(* IEC 61131-3 sources: llm-plc-st-eval/codesys, 25 files *)

(* ---- PRG_Test_A1.st ---- *)
(*
    BANCO DE PRUEBA AUTOVERIFICABLE - Tarea A1 (FB_PID con anti-windup por clamping)
    ---------------------------------------------------------------------------
    Validado en codesys/validar_harness_A1.py: 12 implementaciones (3 correctas,
    con integracion rectangular, integral previa y trapezoidal, y 9 defectuosas).
    Tabla generada desde el validador. tipo: 0 = valor +-tol, 1 = CV <= eVal,
    2 = CV >= eVal.

    TOLERANCIAS (aprobadas por Luis y su asesora, 30-09-2026):
  solo P: +-0.01 | integral: +-2 pasos de muestreo | derivada: +-5 % del termino
  derivativo | saturacion exacta (+-0.001) | anti-windup: sale de la saturacion en
  menos de 1 s tras invertir el error | sentido: PV < SP -> CV sube.

TIEMPO VIRTUAL: ciclo := T#100MS fijo; pasos por NUMERO DE LLAMADAS. Cada
escenario usa su PROPIA instancia del FB (fbP, fbI, fbD, fbW), para que el estado
interno de un escenario (p. ej. una integral acumulada) no contamine otro.

Paso  instancia  (Kp, Ti, Td, SP, PV) llamadas -> comprobacion
  0   fbP  (2, 0, 0, 50, 40)     5 -> CV = 20.0 +-0.01     solo P, sentido
  1   fbP  (2, 0, 0, 50, 60)     5 -> CV = 0.0 +-0.001     saturacion baja
  2   fbP  (2, 0, 0, 50,-20)     5 -> CV = 100.0 +-0.001   saturacion alta
  3   fbP  (2,-1, 0, 50, 45)     5 -> CV = 10.0 +-0.01     Ti < 0: sin integral
  4   fbI  (1,10, 0, 50, 45)   100 -> CV = 10.0 +-0.10     5 + 0.5*10 s
  5   fbI  (1,10, 0, 50, 45)   100 -> CV = 15.0 +-0.10     5 + 0.5*20 s
  6   fbD  (1, 0, 2, 50+0.1k, 40) 50 -> CV = 17.0 +-0.10   e = 15, Td*de/dt = 2 (SP en rampa:
                                                           la derivada sobre PV daria 0)
  7   fbW  (1, 5, 0,100,  0)   300 -> CV = 100.0 +-0.001   30 s saturado en alto
  8   fbW  (1, 5, 0,100,110)    10 -> CV <= 99.5            sale de 100 en < 1 s
  9   fbW  (1, 5, 0,  0,200)   300 -> CV = 0.0 +-0.001     30 s saturado en bajo
 10   fbW  (1, 5, 0,  0,-10)    10 -> CV >= 0.5             sale de 0 en < 1 s
*)
PROGRAM PRG_Test_A1
VAR CONSTANT
    ULTIMO_PASO : INT := 10;
END_VAR
VAR
    fbP, fbI, fbD, fbW : FB_PID;    (* una instancia por escenario *)
    ins        : INT;
    Kp, Ti, Td : REAL;
    SPbase, PV : REAL;
    rampa      : BOOL;
    kRampa     : INT;
    SP, CV     : REAL;
    nLlamadas, k, tipo : INT;
    eVal, tol  : REAL;
    bien       : BOOL;
    paso       : INT := 0;
    finalizado : BOOL;

    resultado : ARRAY[0..10] OF INT;
    nPasan    : INT;
    veredicto : INT := 0;
    i         : INT;
END_VAR

IF NOT finalizado THEN
    (* 1. Definicion del paso *)
    CASE paso OF
        0: ins := 0; Kp := 2.0; Ti := 0.0; Td := 0.0; SPbase := 50.0; rampa := FALSE; PV := 40.0; nLlamadas := 5; tipo := 0; eVal := 20.0; tol := 0.01;
        1: ins := 0; Kp := 2.0; Ti := 0.0; Td := 0.0; SPbase := 50.0; rampa := FALSE; PV := 60.0; nLlamadas := 5; tipo := 0; eVal := 0.0; tol := 0.001;
        2: ins := 0; Kp := 2.0; Ti := 0.0; Td := 0.0; SPbase := 50.0; rampa := FALSE; PV := -20.0; nLlamadas := 5; tipo := 0; eVal := 100.0; tol := 0.001;
        3: ins := 0; Kp := 2.0; Ti := -1.0; Td := 0.0; SPbase := 50.0; rampa := FALSE; PV := 45.0; nLlamadas := 5; tipo := 0; eVal := 10.0; tol := 0.01;
        4: ins := 1; Kp := 1.0; Ti := 10.0; Td := 0.0; SPbase := 50.0; rampa := FALSE; PV := 45.0; nLlamadas := 100; tipo := 0; eVal := 10.0; tol := 0.1;
        5: ins := 1; Kp := 1.0; Ti := 10.0; Td := 0.0; SPbase := 50.0; rampa := FALSE; PV := 45.0; nLlamadas := 100; tipo := 0; eVal := 15.0; tol := 0.1;
        6: ins := 2; Kp := 1.0; Ti := 0.0; Td := 2.0; SPbase := 50.0; rampa := TRUE; PV := 40.0; nLlamadas := 50; tipo := 0; eVal := 17.0; tol := 0.1;
        7: ins := 3; Kp := 1.0; Ti := 5.0; Td := 0.0; SPbase := 100.0; rampa := FALSE; PV := 0.0; nLlamadas := 300; tipo := 0; eVal := 100.0; tol := 0.001;
        8: ins := 3; Kp := 1.0; Ti := 5.0; Td := 0.0; SPbase := 100.0; rampa := FALSE; PV := 110.0; nLlamadas := 10; tipo := 1; eVal := 99.5; tol := 0.0;
        9: ins := 3; Kp := 1.0; Ti := 5.0; Td := 0.0; SPbase := 0.0; rampa := FALSE; PV := 200.0; nLlamadas := 300; tipo := 0; eVal := 0.0; tol := 0.001;
        10: ins := 3; Kp := 1.0; Ti := 5.0; Td := 0.0; SPbase := 0.0; rampa := FALSE; PV := -10.0; nLlamadas := 10; tipo := 2; eVal := 0.5; tol := 0.0;
    END_CASE

    (* 2. Consigna (en rampa en el escenario derivativo) *)
    IF rampa THEN
        kRampa := kRampa + 1;
        SP := SPbase + 0.1 * INT_TO_REAL(kRampa);
    ELSE
        SP := SPbase;
    END_IF

    (* 3. Una llamada por scan a la instancia del escenario, ciclo virtual 100 ms *)
    CASE ins OF
        0: fbP(SP := SP, PV := PV, Kp := Kp, Ti := Ti, Td := Td, ciclo := T#100MS); CV := fbP.CV;
        1: fbI(SP := SP, PV := PV, Kp := Kp, Ti := Ti, Td := Td, ciclo := T#100MS); CV := fbI.CV;
        2: fbD(SP := SP, PV := PV, Kp := Kp, Ti := Ti, Td := Td, ciclo := T#100MS); CV := fbD.CV;
        3: fbW(SP := SP, PV := PV, Kp := Kp, Ti := Ti, Td := Td, ciclo := T#100MS); CV := fbW.CV;
    END_CASE
    k := k + 1;

    (* 4. Evaluacion al completar las llamadas del paso *)
    IF k >= nLlamadas THEN
        CASE tipo OF
            0: bien := ABS(CV - eVal) <= tol;
            1: bien := CV <= eVal;
            2: bien := CV >= eVal;
        END_CASE
        IF bien THEN
            resultado[paso] := 1;
        ELSE
            resultado[paso] := 2;
        END_IF
        k := 0;
        IF paso < ULTIMO_PASO THEN
            paso := paso + 1;
        ELSE
            finalizado := TRUE;
        END_IF
    END_IF
END_IF

(* 5. Veredicto global *)
IF finalizado AND veredicto = 0 THEN
    nPasan := 0;
    FOR i := 0 TO ULTIMO_PASO DO
        IF resultado[i] = 1 THEN
            nPasan := nPasan + 1;
        END_IF
    END_FOR
    IF nPasan = (ULTIMO_PASO + 1) THEN
        veredicto := 1;
    ELSE
        veredicto := 2;
    END_IF
END_IF

(* ---- PRG_Test_A2.st ---- *)
(*
    BANCO DE PRUEBA AUTOVERIFICABLE - Tarea A2 (FB_Batch: receta por lotes de 5 fases)
    ---------------------------------------------------------------------------
    Validado en codesys/validar_harness_A2.py: 9 implementaciones (1 correcta y
    8 defectuosas), ciclos de 4, 10 y 20 ms. Tabla generada desde el validador.
    Al final de cada paso se exige la fase esperada y que este activa exactamente
    la salida de esa fase (fase 0: ninguna).

    Paso: (nA,nB,nVac,ini,abo,temp) duracion -> fase esperada
  0 (F,F,F,F,F,20)   0.2 s -> 0   reposo CON producto
  1 (F,F,F,F,T,20)   0.2 s -> 0   abort en reposo: sin efecto
  2 (F,F,F,T,F,20)   0.2 s -> 1   inicio
  3 (F,F,F,F,F,20)   0.2 s -> 1   espera nivelA
  4 (T,F,F,F,F,20)   0.2 s -> 2
  5 (T,F,F,T,F,20)   0.2 s -> 2   inicio durante la receta: se ignora
  6 (T,T,F,F,F,20)   0.2 s -> 3
  7 (T,T,F,F,F,59.9) 0.2 s -> 3   59.9 no basta
  8 (T,T,F,F,F,60.0) 0.2 s -> 4   60.0 o mas
  9 (T,T,F,F,F,60.0) 118  s -> 4   mezcla: aun no cumple 120 s
 10 (T,T,F,F,F,60.0) 3.0 s -> 5   ya cumplio
 11 (T,T,T,F,F,60.0) 0.2 s -> 0   vacio: reposo
 12 (F,F,F,T,F,20)   0.2 s -> 1   nueva receta (con producto)
 13 (F,F,F,F,T,20)   0.2 s -> 5   abort con producto: descarga
 14 (F,F,F,F,F,20)   0.2 s -> 5   sigue descargando
 15 (F,F,T,F,F,20)   0.2 s -> 0
 16 (F,F,T,T,F,20)   0.2 s -> 1   receta con reactor vacio
 17 (F,F,T,F,T,20)   0.2 s -> 0   abort sin producto: directo a reposo
 18 (F,F,F,T,F,20)   0.2 s -> 1
 19 (T,F,F,F,F,20)   0.2 s -> 2
 20 (T,T,F,F,F,20)   0.2 s -> 3   calentando
 21 (T,T,F,F,T,20)   0.2 s -> 5   abort en fase 3: calentador cerrado, descarga
 22 (T,T,F,F,F,20)   0.2 s -> 5
 23 (T,T,F,F,T,20)   0.2 s -> 5   abort durante la descarga: continua
 24 (T,T,T,F,F,20)   0.2 s -> 0
*)
PROGRAM PRG_Test_A2
VAR CONSTANT
    ULTIMO_PASO : INT := 24;
END_VAR
VAR
    fb : FB_Batch;                  (* bloque bajo prueba *)
    nivelA, nivelB, nivelVacio, btnInicio, btnAbort : BOOL;
    temp  : REAL;
    eFase : INT;
    salidasOk : BOOL;

    paso       : INT := 0;
    tEspera    : TIME;
    tPaso      : TON;
    pulsoReset : BOOL;
    finalizado : BOOL;

    resultado : ARRAY[0..24] OF INT;
    nPasan    : INT;
    veredicto : INT := 0;
    i         : INT;
END_VAR

(* 1. Entradas, duracion y fase esperada del paso *)
IF NOT finalizado THEN
    CASE paso OF
        0: nivelA := FALSE; nivelB := FALSE; nivelVacio := FALSE; btnInicio := FALSE; btnAbort := FALSE;
            temp := 20.0; tEspera := T#200MS; eFase := 0;
        1: nivelA := FALSE; nivelB := FALSE; nivelVacio := FALSE; btnInicio := FALSE; btnAbort := TRUE;
            temp := 20.0; tEspera := T#200MS; eFase := 0;
        2: nivelA := FALSE; nivelB := FALSE; nivelVacio := FALSE; btnInicio := TRUE; btnAbort := FALSE;
            temp := 20.0; tEspera := T#200MS; eFase := 1;
        3: nivelA := FALSE; nivelB := FALSE; nivelVacio := FALSE; btnInicio := FALSE; btnAbort := FALSE;
            temp := 20.0; tEspera := T#200MS; eFase := 1;
        4: nivelA := TRUE; nivelB := FALSE; nivelVacio := FALSE; btnInicio := FALSE; btnAbort := FALSE;
            temp := 20.0; tEspera := T#200MS; eFase := 2;
        5: nivelA := TRUE; nivelB := FALSE; nivelVacio := FALSE; btnInicio := TRUE; btnAbort := FALSE;
            temp := 20.0; tEspera := T#200MS; eFase := 2;
        6: nivelA := TRUE; nivelB := TRUE; nivelVacio := FALSE; btnInicio := FALSE; btnAbort := FALSE;
            temp := 20.0; tEspera := T#200MS; eFase := 3;
        7: nivelA := TRUE; nivelB := TRUE; nivelVacio := FALSE; btnInicio := FALSE; btnAbort := FALSE;
            temp := 59.9; tEspera := T#200MS; eFase := 3;
        8: nivelA := TRUE; nivelB := TRUE; nivelVacio := FALSE; btnInicio := FALSE; btnAbort := FALSE;
            temp := 60.0; tEspera := T#200MS; eFase := 4;
        9: nivelA := TRUE; nivelB := TRUE; nivelVacio := FALSE; btnInicio := FALSE; btnAbort := FALSE;
            temp := 60.0; tEspera := T#118000MS; eFase := 4;
        10: nivelA := TRUE; nivelB := TRUE; nivelVacio := FALSE; btnInicio := FALSE; btnAbort := FALSE;
            temp := 60.0; tEspera := T#3000MS; eFase := 5;
        11: nivelA := TRUE; nivelB := TRUE; nivelVacio := TRUE; btnInicio := FALSE; btnAbort := FALSE;
            temp := 60.0; tEspera := T#200MS; eFase := 0;
        12: nivelA := FALSE; nivelB := FALSE; nivelVacio := FALSE; btnInicio := TRUE; btnAbort := FALSE;
            temp := 20.0; tEspera := T#200MS; eFase := 1;
        13: nivelA := FALSE; nivelB := FALSE; nivelVacio := FALSE; btnInicio := FALSE; btnAbort := TRUE;
            temp := 20.0; tEspera := T#200MS; eFase := 5;
        14: nivelA := FALSE; nivelB := FALSE; nivelVacio := FALSE; btnInicio := FALSE; btnAbort := FALSE;
            temp := 20.0; tEspera := T#200MS; eFase := 5;
        15: nivelA := FALSE; nivelB := FALSE; nivelVacio := TRUE; btnInicio := FALSE; btnAbort := FALSE;
            temp := 20.0; tEspera := T#200MS; eFase := 0;
        16: nivelA := FALSE; nivelB := FALSE; nivelVacio := TRUE; btnInicio := TRUE; btnAbort := FALSE;
            temp := 20.0; tEspera := T#200MS; eFase := 1;
        17: nivelA := FALSE; nivelB := FALSE; nivelVacio := TRUE; btnInicio := FALSE; btnAbort := TRUE;
            temp := 20.0; tEspera := T#200MS; eFase := 0;
        18: nivelA := FALSE; nivelB := FALSE; nivelVacio := FALSE; btnInicio := TRUE; btnAbort := FALSE;
            temp := 20.0; tEspera := T#200MS; eFase := 1;
        19: nivelA := TRUE; nivelB := FALSE; nivelVacio := FALSE; btnInicio := FALSE; btnAbort := FALSE;
            temp := 20.0; tEspera := T#200MS; eFase := 2;
        20: nivelA := TRUE; nivelB := TRUE; nivelVacio := FALSE; btnInicio := FALSE; btnAbort := FALSE;
            temp := 20.0; tEspera := T#200MS; eFase := 3;
        21: nivelA := TRUE; nivelB := TRUE; nivelVacio := FALSE; btnInicio := FALSE; btnAbort := TRUE;
            temp := 20.0; tEspera := T#200MS; eFase := 5;
        22: nivelA := TRUE; nivelB := TRUE; nivelVacio := FALSE; btnInicio := FALSE; btnAbort := FALSE;
            temp := 20.0; tEspera := T#200MS; eFase := 5;
        23: nivelA := TRUE; nivelB := TRUE; nivelVacio := FALSE; btnInicio := FALSE; btnAbort := TRUE;
            temp := 20.0; tEspera := T#200MS; eFase := 5;
        24: nivelA := TRUE; nivelB := TRUE; nivelVacio := TRUE; btnInicio := FALSE; btnAbort := FALSE;
            temp := 20.0; tEspera := T#200MS; eFase := 0;
    END_CASE
END_IF

(* 2. Asentamiento del paso *)
tPaso(IN := NOT pulsoReset, PT := tEspera);
pulsoReset := FALSE;

(* 3. Bloque bajo prueba *)
fb(nivelA := nivelA, nivelB := nivelB, nivelVacio := nivelVacio, btnInicio := btnInicio,
   btnAbort := btnAbort, temp := temp);

(* 4. Evaluacion: fase y exactamente la salida de esa fase *)
IF tPaso.Q AND NOT finalizado THEN
    salidasOk := (fb.vA = (eFase = 1)) AND (fb.vB = (eFase = 2)) AND (fb.calentador = (eFase = 3))
                 AND (fb.mezclador = (eFase = 4)) AND (fb.vDescarga = (eFase = 5));
    IF (fb.fase = eFase) AND salidasOk THEN
        resultado[paso] := 1;
    ELSE
        resultado[paso] := 2;
    END_IF
    pulsoReset := TRUE;
    IF paso < ULTIMO_PASO THEN
        paso := paso + 1;
    ELSE
        finalizado := TRUE;
    END_IF
END_IF

(* 5. Veredicto global *)
IF finalizado AND veredicto = 0 THEN
    nPasan := 0;
    FOR i := 0 TO ULTIMO_PASO DO
        IF resultado[i] = 1 THEN
            nPasan := nPasan + 1;
        END_IF
    END_FOR
    IF nPasan = (ULTIMO_PASO + 1) THEN
        veredicto := 1;
    ELSE
        veredicto := 2;
    END_IF
END_IF

(* ---- PRG_Test_A3.st ---- *)
(*
    BANCO DE PRUEBA AUTOVERIFICABLE - Tarea A3 (FB_Com: peticion/respuesta con reintentos)
    ---------------------------------------------------------------------------
    Validado en codesys/validar_harness_A3.py: 9 implementaciones (1 correcta y
    8 defectuosas), ciclos de 4, 10 y 20 ms. Tabla generada desde el validador.
    rxOk se aplica como pulso de UN scan al entrar en el paso (ver validador).
    eN = -1 o eTx = -1: ese valor no se evalua en el paso.

    Paso: (txReq, pulso rxOk, rxData) duracion -> (ocupado, ok, error, nIntentos, txData)   [- = no se evalua]
  0 (F,-,0)   0.20 s -> (F,F,F,-,-)  reposo
  1 (T,-,0)   0.20 s -> (T,F,F,1,100) flanco: intento 1
  2 (F,-,0)   0.20 s -> (T,F,F,1,-)   0.40 s: aun intento 1   (plazo corto)
  3 (F,-,0)   0.25 s -> (T,F,F,2,-)   0.65 s: intento 2        (plazo largo / sin reintento)
  4 (F,P,100) 0.20 s -> (F,T,F,2,-)   eco correcto: ok, conserva nIntentos=2
  5 (F,-,0)   0.30 s -> (F,T,F,2,-)   ok permanece
  6 (T,-,0)   0.10 s -> (T,F,F,1,100) nuevo intercambio: ok se borra
  7 (F,P,55)  0.10 s -> (T,F,F,2,-)   eco erroneo: falla el intento 1
  8 (T,-,0)   0.10 s -> (T,F,F,2,-)   flanco de txReq durante el intercambio: se ignora
  9 (T,-,0)   0.50 s -> (T,F,F,3,-)   vence el intento 2
 10 (T,-,0)   0.40 s -> (F,F,T,3,-)   vence el intento 3: error
 11 (F,-,0)   0.30 s -> (F,F,T,3,-)   error permanece, nIntentos se conserva
 12 (T,-,0)   0.20 s -> (T,F,F,1,100) nuevo intercambio: error se borra
 13 (T,-,0)   0.20 s -> (T,F,F,1,-)   ~0.41-0.46 s del intento 1 (segun el ciclo)
 14 (T,P,100) 0.20 s -> (F,T,F,1,-)   eco al inicio del paso: dentro del plazo (plazo demasiado corto)
NOTA: la primera version usaba 0.25 s en el paso 13 y REPROBABA a la correcta con
ciclo de 20 ms (el eco llegaba a ~0.51 s): cada cambio de paso consume un scan.
*)
PROGRAM PRG_Test_A3
VAR CONSTANT
    ULTIMO_PASO : INT := 14;
END_VAR
VAR
    fb : FB_Com;                    (* bloque bajo prueba *)
    txReq, rxOk : BOOL;
    rxData      : INT;
    pulsoStep   : BOOL;             (* el paso aplica un pulso de rxOk *)
    pendiente   : BOOL;
    pasoCargado : INT := -1;
    eOcup, eOk, eErr : BOOL;
    eN, eTx     : INT;

    paso       : INT := 0;
    tEspera    : TIME;
    tPaso      : TON;
    pulsoReset : BOOL;
    finalizado : BOOL;

    resultado : ARRAY[0..14] OF INT;
    nPasan    : INT;
    veredicto : INT := 0;
    i         : INT;
END_VAR

(* 1. Entradas, duracion y valores esperados del paso *)
IF NOT finalizado THEN
    CASE paso OF
        0: txReq := FALSE; pulsoStep := FALSE; rxData := 0; tEspera := T#200MS;
            eOcup := FALSE; eOk := FALSE; eErr := FALSE; eN := -1; eTx := -1;
        1: txReq := TRUE; pulsoStep := FALSE; rxData := 0; tEspera := T#200MS;
            eOcup := TRUE; eOk := FALSE; eErr := FALSE; eN := 1; eTx := 100;
        2: txReq := FALSE; pulsoStep := FALSE; rxData := 0; tEspera := T#200MS;
            eOcup := TRUE; eOk := FALSE; eErr := FALSE; eN := 1; eTx := -1;
        3: txReq := FALSE; pulsoStep := FALSE; rxData := 0; tEspera := T#250MS;
            eOcup := TRUE; eOk := FALSE; eErr := FALSE; eN := 2; eTx := -1;
        4: txReq := FALSE; pulsoStep := TRUE; rxData := 100; tEspera := T#200MS;
            eOcup := FALSE; eOk := TRUE; eErr := FALSE; eN := 2; eTx := -1;
        5: txReq := FALSE; pulsoStep := FALSE; rxData := 0; tEspera := T#300MS;
            eOcup := FALSE; eOk := TRUE; eErr := FALSE; eN := 2; eTx := -1;
        6: txReq := TRUE; pulsoStep := FALSE; rxData := 0; tEspera := T#100MS;
            eOcup := TRUE; eOk := FALSE; eErr := FALSE; eN := 1; eTx := 100;
        7: txReq := FALSE; pulsoStep := TRUE; rxData := 55; tEspera := T#100MS;
            eOcup := TRUE; eOk := FALSE; eErr := FALSE; eN := 2; eTx := -1;
        8: txReq := TRUE; pulsoStep := FALSE; rxData := 0; tEspera := T#100MS;
            eOcup := TRUE; eOk := FALSE; eErr := FALSE; eN := 2; eTx := -1;
        9: txReq := TRUE; pulsoStep := FALSE; rxData := 0; tEspera := T#500MS;
            eOcup := TRUE; eOk := FALSE; eErr := FALSE; eN := 3; eTx := -1;
        10: txReq := TRUE; pulsoStep := FALSE; rxData := 0; tEspera := T#400MS;
            eOcup := FALSE; eOk := FALSE; eErr := TRUE; eN := 3; eTx := -1;
        11: txReq := FALSE; pulsoStep := FALSE; rxData := 0; tEspera := T#300MS;
            eOcup := FALSE; eOk := FALSE; eErr := TRUE; eN := 3; eTx := -1;
        12: txReq := TRUE; pulsoStep := FALSE; rxData := 0; tEspera := T#200MS;
            eOcup := TRUE; eOk := FALSE; eErr := FALSE; eN := 1; eTx := 100;
        13: txReq := TRUE; pulsoStep := FALSE; rxData := 0; tEspera := T#200MS;
            eOcup := TRUE; eOk := FALSE; eErr := FALSE; eN := 1; eTx := -1;
        14: txReq := TRUE; pulsoStep := TRUE; rxData := 100; tEspera := T#200MS;
            eOcup := FALSE; eOk := TRUE; eErr := FALSE; eN := 1; eTx := -1;
    END_CASE
END_IF

(* 2. Pulso de rxOk de un solo scan al entrar en el paso *)
IF paso <> pasoCargado THEN
    pendiente := pulsoStep;
    pasoCargado := paso;
END_IF
rxOk := pendiente AND NOT finalizado;
pendiente := FALSE;

(* 3. Asentamiento del paso *)
tPaso(IN := NOT pulsoReset, PT := tEspera);
pulsoReset := FALSE;

(* 4. Bloque bajo prueba *)
fb(txReq := txReq, rxOk := rxOk, rxData := rxData);

(* 5. Evaluacion *)
IF tPaso.Q AND NOT finalizado THEN
    IF (fb.ocupado = eOcup) AND (fb.ok = eOk) AND (fb.error = eErr)
       AND ((eN < 0) OR (fb.nIntentos = eN)) AND ((eTx < 0) OR (fb.txData = eTx)) THEN
        resultado[paso] := 1;
    ELSE
        resultado[paso] := 2;
    END_IF
    pulsoReset := TRUE;
    IF paso < ULTIMO_PASO THEN
        paso := paso + 1;
    ELSE
        finalizado := TRUE;
    END_IF
END_IF

(* 6. Veredicto global *)
IF finalizado AND veredicto = 0 THEN
    nPasan := 0;
    FOR i := 0 TO ULTIMO_PASO DO
        IF resultado[i] = 1 THEN
            nPasan := nPasan + 1;
        END_IF
    END_FOR
    IF nPasan = (ULTIMO_PASO + 1) THEN
        veredicto := 1;
    ELSE
        veredicto := 2;
    END_IF
END_IF

(* ---- PRG_Test_A4.st ---- *)
(*
    BANCO DE PRUEBA AUTOVERIFICABLE - Tarea A4 (FB_Rampa: consigna con rampa)
    ---------------------------------------------------------------------------
    Validado en codesys/validar_harness_A4.py: 8 implementaciones (1 correcta y
    7 defectuosas). Tabla generada desde el validador.

    TIEMPO VIRTUAL: se pasa siempre ciclo := T#10MS y cada paso dura un NUMERO DE
    LLAMADAS (una por scan), no un tiempo. El resultado no depende del ciclo real.
    Tolerancia 0.01 en el valor final del paso; vigilancia de sobrepaso con 0.001
    (vig = 1: CVvel <= objetivo; vig = 2: CVvel >= objetivo, en cada llamada).

    Paso: (SP, paro) llamadas -> CVvel esperado   [vigilancia]
  0 (0.05,F)  1 ->  0.05   escalon menor que el incremento (0.1): sin sobrepaso [CV <= 0.05]
  1 ( 0,F)    1 ->  0.0    idem al bajar                                        [CV >= 0]
  2 (50,F)  300 -> 30.0    subida 10 %/s
  3 (50,F)  300 -> 50.0    llega y se queda           [CV <= 50]
  4 (20,F)  100 -> 30.0    bajada 20 %/s
  5 (20,F)  100 -> 20.0                               [CV >= 20]
  6 (80,F)  200 -> 40.0
  7 (80,T)   50 -> 20.0    paro rapido 40 %/s
  8 (80,T)  100 ->  0.0                               [CV >= 0]
  9 (80,T)   50 ->  0.0    permanece en 0 con paro    [CV <= 0]
 10 (80,F)  100 -> 10.0    sin paro: vuelve a subir
 11 (10.05,F) 1 -> 10.05                              [CV <= 10.05]
 12 ( 9,F)   10 ->  9.0                               [CV >= 9]
El sobrepaso se prueba PRIMERO (pasos 0 y 1), desde 0.0 y sin acumulacion previa:
asi el paso de fallo de un bloque que no acota no depende del redondeo de REAL
de 32 bits frente al float de 64 bits del validador.
*)
PROGRAM PRG_Test_A4
VAR CONSTANT
    ULTIMO_PASO : INT  := 12;
    TOL         : REAL := 0.01;
    TOL_VIG     : REAL := 0.001;
END_VAR
VAR
    fb : FB_Rampa;                  (* bloque bajo prueba *)
    SPvel      : REAL;
    paroRapido : BOOL;
    nLlamadas  : INT;               (* llamadas del paso *)
    k          : INT;               (* llamadas hechas en el paso *)
    eCV        : REAL;
    vig        : INT;
    violacion  : BOOL;
    paso       : INT := 0;
    finalizado : BOOL;

    resultado : ARRAY[0..12] OF INT;
    nPasan    : INT;
    veredicto : INT := 0;
    i         : INT;
END_VAR

IF NOT finalizado THEN
    (* 1. Definicion del paso *)
    CASE paso OF
        0: SPvel := 0.05; paroRapido := FALSE; nLlamadas := 1; eCV := 0.05; vig := 1;
        1: SPvel := 0.0; paroRapido := FALSE; nLlamadas := 1; eCV := 0.0; vig := 2;
        2: SPvel := 50.0; paroRapido := FALSE; nLlamadas := 300; eCV := 30.0; vig := 0;
        3: SPvel := 50.0; paroRapido := FALSE; nLlamadas := 300; eCV := 50.0; vig := 1;
        4: SPvel := 20.0; paroRapido := FALSE; nLlamadas := 100; eCV := 30.0; vig := 0;
        5: SPvel := 20.0; paroRapido := FALSE; nLlamadas := 100; eCV := 20.0; vig := 2;
        6: SPvel := 80.0; paroRapido := FALSE; nLlamadas := 200; eCV := 40.0; vig := 0;
        7: SPvel := 80.0; paroRapido := TRUE; nLlamadas := 50; eCV := 20.0; vig := 0;
        8: SPvel := 80.0; paroRapido := TRUE; nLlamadas := 100; eCV := 0.0; vig := 2;
        9: SPvel := 80.0; paroRapido := TRUE; nLlamadas := 50; eCV := 0.0; vig := 1;
        10: SPvel := 80.0; paroRapido := FALSE; nLlamadas := 100; eCV := 10.0; vig := 0;
        11: SPvel := 10.05; paroRapido := FALSE; nLlamadas := 1; eCV := 10.05; vig := 1;
        12: SPvel := 9.0; paroRapido := FALSE; nLlamadas := 10; eCV := 9.0; vig := 2;
    END_CASE

    (* 2. Una llamada por scan con ciclo virtual de 10 ms *)
    fb(SPvel := SPvel, paroRapido := paroRapido, ciclo := T#10MS);
    k := k + 1;

    (* 3. Vigilancia de sobrepaso *)
    IF ((vig = 1) AND (fb.CVvel > eCV + TOL_VIG)) OR ((vig = 2) AND (fb.CVvel < eCV - TOL_VIG)) THEN
        violacion := TRUE;
    END_IF

    (* 4. Evaluacion al completar las llamadas del paso *)
    IF k >= nLlamadas THEN
        IF (ABS(fb.CVvel - eCV) <= TOL) AND NOT violacion THEN
            resultado[paso] := 1;
        ELSE
            resultado[paso] := 2;
        END_IF
        k := 0;
        violacion := FALSE;
        IF paso < ULTIMO_PASO THEN
            paso := paso + 1;
        ELSE
            finalizado := TRUE;
        END_IF
    END_IF
END_IF

(* 5. Veredicto global *)
IF finalizado AND veredicto = 0 THEN
    nPasan := 0;
    FOR i := 0 TO ULTIMO_PASO DO
        IF resultado[i] = 1 THEN
            nPasan := nPasan + 1;
        END_IF
    END_FOR
    IF nPasan = (ULTIMO_PASO + 1) THEN
        veredicto := 1;
    ELSE
        veredicto := 2;
    END_IF
END_IF

(* ---- PRG_Test_A5.st ---- *)
(*
    BANCO DE PRUEBA AUTOVERIFICABLE - Tarea A5 (FB_Registro: buffer circular de eventos)
    ---------------------------------------------------------------------------
    Validado en codesys/validar_harness_A5.py: 9 implementaciones (2 correctas,
    que acumulan el tiempo antes y despues de registrar, y 7 defectuosas).
    Tabla generada desde el validador.
    TIEMPO VIRTUAL: ciclo := T#10MS fijo; pasos por numero de llamadas (una por
    scan). Para el ultimo evento se acepta marca = g*10 ms o (g-1)*10 ms.
    pM/p2 = -1: no se comprueba contenido en ese paso.

    Paso: llamadas/eventos -> (indice, nEventos, comprobacion de contenido)
  0 5 llamadas sin evento ..................... (-1, 0)
  1 evento 11 con nuevoEvento sostenido 3 llamadas (0, 1)  buffer[0]=11 + marca
  2 2 llamadas sin flanco ..................... (0, 1)
  3 19 eventos (12..30) ....................... (19, 20) buffer[19]=30 + marca; buffer[0]=11
  4 1 evento (31): sobrescribe el mas antiguo . (0, 20)  buffer[0]=31 + marca; buffer[1]=12
  5 2 eventos (32, 33) ........................ (2, 20)  buffer[2]=33 + marca; buffer[3]=14
*)
PROGRAM PRG_Test_A5
VAR CONSTANT
    ULTIMO_PASO : INT := 5;
END_VAR
VAR
    fb : FB_Registro;               (* bloque bajo prueba *)
    evento      : INT;
    nuevoEvento : BOOL;
    prevNuevo   : BOOL;
    nEv, libres, sost, cod0 : INT;  (* definicion del paso *)
    eIdx, eN, pM, cM, p2, c2 : INT; (* comprobaciones del paso *)
    L, k        : INT;              (* llamadas del paso / hechas *)
    g, gUlt     : DINT;             (* llamadas totales / del ultimo flanco *)
    bien        : BOOL;
    paso        : INT := 0;
    finalizado  : BOOL;

    resultado : ARRAY[0..5] OF INT;
    nPasan    : INT;
    veredicto : INT := 0;
    i         : INT;
END_VAR

IF NOT finalizado THEN
    (* 1. Definicion del paso *)
    CASE paso OF
        0: nEv := 0; libres := 5; sost := 0; cod0 := 0; eIdx := -1; eN := 0; pM := -1; cM := 0; p2 := -1; c2 := 0;
        1: nEv := 1; libres := 0; sost := 3; cod0 := 11; eIdx := 0; eN := 1; pM := 0; cM := 11; p2 := -1; c2 := 0;
        2: nEv := 0; libres := 2; sost := 0; cod0 := 0; eIdx := 0; eN := 1; pM := -1; cM := 0; p2 := -1; c2 := 0;
        3: nEv := 19; libres := 0; sost := 0; cod0 := 12; eIdx := 19; eN := 20; pM := 19; cM := 30; p2 := 0; c2 := 11;
        4: nEv := 1; libres := 0; sost := 0; cod0 := 31; eIdx := 0; eN := 20; pM := 0; cM := 31; p2 := 1; c2 := 12;
        5: nEv := 2; libres := 0; sost := 0; cod0 := 32; eIdx := 2; eN := 20; pM := 2; cM := 33; p2 := 3; c2 := 14;
    END_CASE
    IF sost > 0 THEN
        L := sost + libres;
    ELSE
        L := 2 * nEv + libres;
    END_IF

    (* 2. Entradas de esta llamada *)
    IF sost > 0 THEN
        IF k < sost THEN
            evento := cod0; nuevoEvento := TRUE;
        ELSE
            evento := 0; nuevoEvento := FALSE;
        END_IF
    ELSIF k < 2 * nEv THEN
        evento := cod0 + k / 2;
        nuevoEvento := (k MOD 2) = 0;
    ELSE
        evento := 0; nuevoEvento := FALSE;
    END_IF

    (* 3. Llamada con ciclo virtual de 10 ms *)
    g := g + 1;
    fb(evento := evento, nuevoEvento := nuevoEvento, ciclo := T#10MS);
    IF nuevoEvento AND NOT prevNuevo THEN
        gUlt := g;
    END_IF
    prevNuevo := nuevoEvento;
    k := k + 1;

    (* 4. Evaluacion al completar el paso *)
    IF k >= L THEN
        bien := (fb.indice = eIdx) AND (fb.nEventos = eN);
        IF pM >= 0 THEN
            bien := bien AND (fb.buffer[pM].codigo = cM)
                    AND ((fb.buffer[pM].marca = DINT_TO_TIME(gUlt * 10)) OR (fb.buffer[pM].marca = DINT_TO_TIME((gUlt - 1) * 10)));
        END_IF
        IF p2 >= 0 THEN
            bien := bien AND (fb.buffer[p2].codigo = c2);
        END_IF
        IF bien THEN
            resultado[paso] := 1;
        ELSE
            resultado[paso] := 2;
        END_IF
        k := 0;
        IF paso < ULTIMO_PASO THEN
            paso := paso + 1;
        ELSE
            finalizado := TRUE;
        END_IF
    END_IF
END_IF

(* 5. Veredicto global *)
IF finalizado AND veredicto = 0 THEN
    nPasan := 0;
    FOR i := 0 TO ULTIMO_PASO DO
        IF resultado[i] = 1 THEN
            nPasan := nPasan + 1;
        END_IF
    END_FOR
    IF nPasan = (ULTIMO_PASO + 1) THEN
        veredicto := 1;
    ELSE
        veredicto := 2;
    END_IF
END_IF

(* ---- PRG_Test_A6.st ---- *)
(*
    BANCO DE PRUEBA AUTOVERIFICABLE - Tarea A6 (FB_Modos: modos jerarquicos con forzado)
    ---------------------------------------------------------------------------
    Validado en codesys/validar_harness_A6.py: 10 implementaciones (1 correcta y
    9 defectuosas), ciclos de 4, 10 y 20 ms. Tabla generada desde el validador.
    Los patrones de 8 bits se codifican como mascara WORD: bit i = elemento [i].
    cmdManual es siempre M = 11001100 (mascara MASK_MANUAL). confirmarForzado se
    aplica como pulso de UN scan al entrar en el paso.

    Paso: (selector, seguro, cmdAuto, idx, val, pulso) -> (modo, actuadores)
  0 (0,F,A, 0,F,-) -> (1, M)        arranca en manual; sin seguro no cambia
  1 (0,F,A, 0,F,-) -> (1, M)
  2 (0,T,A, 0,F,-) -> (0, A)        el cambio pendiente se aplica al activarse seguro
  3 (5,T,A, 0,F,-) -> (0, A)        fuera de rango: se ignora
  4 (-1,T,A,0,F,-) -> (0, A)
  5 (0,T,A2,0,F,-) -> (0, A2)       sigue a cmdAuto
  6 (2,T,A2,0,F,-) -> (2, 00000000) mantenimiento: todo apagado
  7 (2,T,A2,3,T,P) -> (2, 00010000) fuerza actuador[3]
  8 (2,T,A2,8,T,P) -> (2, 00010000) idx fuera de rango: se ignora
  9 (2,T,A2,5,T,P) -> (2, 00010100)
 10 (2,T,A2,3,F,P) -> (2, 00000100) forzado a FALSE
 11 (2,F,A2,0,F,-) -> (2, 00000000) pierde seguro: anula forzados
 12 (2,T,A2,0,F,-) -> (2, 00000000) vuelve el seguro: siguen anulados
 13 (2,T,A2,0,T,P) -> (2, 10000000)
 14 (1,T,A2,0,F,-) -> (1, M)        sale a manual
 15 (2,T,A2,0,F,-) -> (2, 00000000) los forzados de antes no reaparecen
 16 (0,T,A2,0,F,-) -> (0, A2)
*)
PROGRAM PRG_Test_A6
VAR CONSTANT
    ULTIMO_PASO : INT  := 16;
    T_PASO      : TIME := T#100MS;
    MASK_MANUAL : WORD := 51;
END_VAR
VAR
    fb : FB_Modos;                  (* bloque bajo prueba *)
    selector     : INT;
    estadoSeguro : BOOL;
    cmdAuto      : ARRAY[0..7] OF BOOL;
    cmdManual    : ARRAY[0..7] OF BOOL;
    idxForzado   : INT;
    valorForzado : BOOL;
    confirmarForzado : BOOL;
    mAuto, eMask, mAct : WORD;
    eModo        : INT;
    pulsoStep, pendiente : BOOL;
    pasoCargado  : INT := -1;
    b            : INT;

    paso       : INT := 0;
    tPaso      : TON;
    pulsoReset : BOOL;
    finalizado : BOOL;

    resultado : ARRAY[0..16] OF INT;
    nPasan    : INT;
    veredicto : INT := 0;
    i         : INT;
END_VAR

(* 1. Definicion del paso *)
IF NOT finalizado THEN
    CASE paso OF
        0: selector := 0; estadoSeguro := FALSE; mAuto := 85; idxForzado := 0; valorForzado := FALSE; pulsoStep := FALSE; eModo := 1; eMask := 51;
        1: selector := 0; estadoSeguro := FALSE; mAuto := 85; idxForzado := 0; valorForzado := FALSE; pulsoStep := FALSE; eModo := 1; eMask := 51;
        2: selector := 0; estadoSeguro := TRUE; mAuto := 85; idxForzado := 0; valorForzado := FALSE; pulsoStep := FALSE; eModo := 0; eMask := 85;
        3: selector := 5; estadoSeguro := TRUE; mAuto := 85; idxForzado := 0; valorForzado := FALSE; pulsoStep := FALSE; eModo := 0; eMask := 85;
        4: selector := -1; estadoSeguro := TRUE; mAuto := 85; idxForzado := 0; valorForzado := FALSE; pulsoStep := FALSE; eModo := 0; eMask := 85;
        5: selector := 0; estadoSeguro := TRUE; mAuto := 102; idxForzado := 0; valorForzado := FALSE; pulsoStep := FALSE; eModo := 0; eMask := 102;
        6: selector := 2; estadoSeguro := TRUE; mAuto := 102; idxForzado := 0; valorForzado := FALSE; pulsoStep := FALSE; eModo := 2; eMask := 0;
        7: selector := 2; estadoSeguro := TRUE; mAuto := 102; idxForzado := 3; valorForzado := TRUE; pulsoStep := TRUE; eModo := 2; eMask := 8;
        8: selector := 2; estadoSeguro := TRUE; mAuto := 102; idxForzado := 8; valorForzado := TRUE; pulsoStep := TRUE; eModo := 2; eMask := 8;
        9: selector := 2; estadoSeguro := TRUE; mAuto := 102; idxForzado := 5; valorForzado := TRUE; pulsoStep := TRUE; eModo := 2; eMask := 40;
        10: selector := 2; estadoSeguro := TRUE; mAuto := 102; idxForzado := 3; valorForzado := FALSE; pulsoStep := TRUE; eModo := 2; eMask := 32;
        11: selector := 2; estadoSeguro := FALSE; mAuto := 102; idxForzado := 0; valorForzado := FALSE; pulsoStep := FALSE; eModo := 2; eMask := 0;
        12: selector := 2; estadoSeguro := TRUE; mAuto := 102; idxForzado := 0; valorForzado := FALSE; pulsoStep := FALSE; eModo := 2; eMask := 0;
        13: selector := 2; estadoSeguro := TRUE; mAuto := 102; idxForzado := 0; valorForzado := TRUE; pulsoStep := TRUE; eModo := 2; eMask := 1;
        14: selector := 1; estadoSeguro := TRUE; mAuto := 102; idxForzado := 0; valorForzado := FALSE; pulsoStep := FALSE; eModo := 1; eMask := 51;
        15: selector := 2; estadoSeguro := TRUE; mAuto := 102; idxForzado := 0; valorForzado := FALSE; pulsoStep := FALSE; eModo := 2; eMask := 0;
        16: selector := 0; estadoSeguro := TRUE; mAuto := 102; idxForzado := 0; valorForzado := FALSE; pulsoStep := FALSE; eModo := 0; eMask := 102;
    END_CASE
END_IF
FOR b := 0 TO 7 DO
    cmdAuto[b] := (SHR(mAuto, b) AND 1) = 1;
    cmdManual[b] := (SHR(MASK_MANUAL, b) AND 1) = 1;
END_FOR

(* 2. Pulso de confirmarForzado de un scan al entrar en el paso *)
IF paso <> pasoCargado THEN
    pendiente := pulsoStep;
    pasoCargado := paso;
END_IF
confirmarForzado := pendiente AND NOT finalizado;
pendiente := FALSE;

(* 3. Asentamiento del paso *)
tPaso(IN := NOT pulsoReset, PT := T_PASO);
pulsoReset := FALSE;

(* 4. Bloque bajo prueba *)
fb(selector := selector, estadoSeguro := estadoSeguro, cmdAuto := cmdAuto, cmdManual := cmdManual,
   idxForzado := idxForzado, valorForzado := valorForzado, confirmarForzado := confirmarForzado);

(* 5. Evaluacion *)
IF tPaso.Q AND NOT finalizado THEN
    mAct := 0;
    FOR b := 0 TO 7 DO
        IF fb.actuador[b] THEN
            mAct := mAct OR SHL(WORD#1, b);
        END_IF
    END_FOR
    IF (fb.modoActivo = eModo) AND (mAct = eMask) THEN
        resultado[paso] := 1;
    ELSE
        resultado[paso] := 2;
    END_IF
    pulsoReset := TRUE;
    IF paso < ULTIMO_PASO THEN
        paso := paso + 1;
    ELSE
        finalizado := TRUE;
    END_IF
END_IF

(* 6. Veredicto global *)
IF finalizado AND veredicto = 0 THEN
    nPasan := 0;
    FOR i := 0 TO ULTIMO_PASO DO
        IF resultado[i] = 1 THEN
            nPasan := nPasan + 1;
        END_IF
    END_FOR
    IF nPasan = (ULTIMO_PASO + 1) THEN
        veredicto := 1;
    ELSE
        veredicto := 2;
    END_IF
END_IF

(* ---- PRG_Test_B1.st ---- *)
(*
    BANCO DE PRUEBA AUTOVERIFICABLE — Tarea B1 (arranque/paro con enclavamiento)
    ---------------------------------------------------------------------------
    Implementa el protocolo de 7 pasos de la ficha de evaluacion de B1 como
    codigo ST. El programa aplica las entradas paso a paso, compara la salida
    del bloque bajo prueba contra el valor esperado y emite un veredicto.

    Ventaja para la investigacion: la verificacion funcional deja de depender
    de que el investigador manipule variables a mano en linea. El mismo
    protocolo se aplica de forma identica a las 24 respuestas de B1, lo que
    elimina la variabilidad del operador. El veredicto queda en una variable
    que el ScriptEngine puede leer, o que puede volcarse a archivo.

    LO QUE NO HACE: no juzga claridad estructural ni mantenibilidad. Esos
    criterios de la rubrica siguen requiriendo lectura humana del codigo.

    USO: crear este PROGRAM en el proyecto, junto al FUNCTION_BLOCK de la
    respuesta a evaluar. Ejecutar en modo Simulacion. Al terminar la secuencia,
    leer 'veredicto': 1 = supera todos los pasos, 2 = falla al menos uno.
    El arreglo 'resultado' indica que paso concreto fallo.
*)

PROGRAM PRG_Test_B1
VAR CONSTANT
    ULTIMO_PASO : INT := 6;          (* 7 pasos: indices 0..6 *)
    T_ASENTAMIENTO : TIME := T#200MS; (* margen por paso; subir si hay temporizadores *)
END_VAR
VAR
    (* --- Bloque bajo prueba: sustituir por la respuesta a evaluar --- *)
    fb : FB_Motor;

    (* --- Entradas manipuladas por el banco --- *)
    btnMarcha : BOOL;
    btnParo   : BOOL;
    btnEmerg  : BOOL;

    (* --- Control de la secuencia --- *)
    paso       : INT := 0;
    esperado   : BOOL;
    tPaso      : TON;
    pulsoReset : BOOL;
    finalizado : BOOL;

    (* --- Resultados: 0 = pendiente, 1 = pasa, 2 = falla --- *)
    resultado : ARRAY[0..6] OF INT;
    nPasan    : INT;
    veredicto : INT := 0;            (* 0 = en curso, 1 = PASA, 2 = FALLA *)
    i         : INT;
END_VAR

(* 1. Temporizador de asentamiento entre pasos *)
tPaso(IN := NOT pulsoReset, PT := T_ASENTAMIENTO);
pulsoReset := FALSE;

(* 2. Aplicacion de entradas y valor esperado segun el paso *)
IF NOT finalizado THEN
    CASE paso OF
        0:  (* Reposo: ninguna entrada activa *)
            btnMarcha := FALSE; btnParo := FALSE; btnEmerg := FALSE;
            esperado  := FALSE;
        1:  (* Arranque con pulso de marcha *)
            btnMarcha := TRUE;
            esperado  := TRUE;
        2:  (* Se suelta la marcha: debe mantenerse (enclavamiento) *)
            btnMarcha := FALSE;
            esperado  := TRUE;
        3:  (* Paro normal *)
            btnParo   := TRUE;
            esperado  := FALSE;
        4:  (* Rearranque tras paro normal *)
            btnParo   := FALSE; btnMarcha := TRUE;
            esperado  := TRUE;
        5:  (* Paro de emergencia *)
            btnEmerg  := TRUE;
            esperado  := FALSE;
        6:  (* Se libera la emergencia con la marcha aun pulsada:
               NO debe rearrancar solo *)
            btnEmerg  := FALSE;
            esperado  := FALSE;
    END_CASE
END_IF

(* 3. Llamada al bloque bajo prueba *)
fb(btnMarcha := btnMarcha, btnParo := btnParo, btnEmerg := btnEmerg);

(* 4. Evaluacion al vencer el tiempo de asentamiento *)
IF tPaso.Q AND NOT finalizado THEN
    IF fb.motorOn = esperado THEN
        resultado[paso] := 1;
    ELSE
        resultado[paso] := 2;
    END_IF

    pulsoReset := TRUE;              (* reinicia el temporizador un ciclo *)

    IF paso < ULTIMO_PASO THEN
        paso := paso + 1;
    ELSE
        finalizado := TRUE;
    END_IF
END_IF

(* 5. Veredicto global *)
IF finalizado AND veredicto = 0 THEN
    nPasan := 0;
    FOR i := 0 TO ULTIMO_PASO DO
        IF resultado[i] = 1 THEN
            nPasan := nPasan + 1;
        END_IF
    END_FOR

    IF nPasan = (ULTIMO_PASO + 1) THEN
        veredicto := 1;              (* supera el protocolo completo *)
    ELSE
        veredicto := 2;              (* falla al menos un paso *)
    END_IF
END_IF

(* ---- PRG_Test_B2.st ---- *)
(*
    BANCO DE PRUEBA AUTOVERIFICABLE — Tarea B2 (valvula con retardo TON de 5 s)
    ---------------------------------------------------------------------------
    PLANTILLA PARA TAREAS CON TEMPORIZADORES.

    Diferencia clave respecto a PRG_Test_B1: el tiempo de asentamiento es
    DISTINTO EN CADA PASO. Un valor fijo corto (200 ms) haria fallar a bloques
    correctos, porque evaluaria la salida antes de que venza el temporizador
    interno del bloque bajo prueba. Con un TON de 5 s, el paso que espera la
    apertura necesita mas de 5 s de asentamiento.

    Usa esta plantilla (y no la de B1) en las tareas B2, B5, B6, I1, I2, I4,
    I5 e I8, que incluyen temporizacion. La de B1 solo sirve para logica
    puramente combinacional o de enclavamiento sin retardos.

    ATENCION AL TIEMPO REAL: la simulacion corre en tiempo real, de modo que
    un banco con esperas de 6 s por paso tarda unos 20 s por respuesta. Para
    24 respuestas de una tarea son unos 8 minutos; asumible. En tareas con
    retardos largos (B5 usa TOF de 30 s; I1 encadena 20+4+15 s) conviene
    estimar el tiempo total antes de lanzar el lote.
*)

PROGRAM PRG_Test_B2
VAR CONSTANT
    ULTIMO_PASO : INT := 5;          (* 6 pasos: indices 0..5 *)
END_VAR
VAR
    (* --- Bloque bajo prueba --- *)
    fb : FB_Valvula;

    (* --- Entrada manipulada por el banco --- *)
    nivelAlto : BOOL;

    (* --- Control de la secuencia --- *)
    paso       : INT := 0;
    esperado   : BOOL;
    tEspera    : TIME;               (* asentamiento del paso en curso *)
    tPaso      : TON;
    pulsoReset : BOOL;
    finalizado : BOOL;

    (* --- Resultados: 0 = pendiente, 1 = pasa, 2 = falla --- *)
    resultado : ARRAY[0..5] OF INT;
    nPasan    : INT;
    veredicto : INT := 0;            (* 0 = en curso, 1 = PASA, 2 = FALLA *)
    i         : INT;
END_VAR

(* 1. Definicion del paso en curso: entrada, espera y valor esperado.
      Se evalua antes del temporizador porque tEspera lo alimenta. *)
IF NOT finalizado THEN
    CASE paso OF
        0:  (* Reposo *)
            nivelAlto := FALSE;
            tEspera   := T#500MS;
            esperado  := FALSE;
        1:  (* Nivel alto durante 3 s: aun NO debe abrir (el TON pide 5 s) *)
            nivelAlto := TRUE;
            tEspera   := T#3S;
            esperado  := FALSE;
        2:  (* Se mantiene 3 s mas (6 s acumulados): ya debe abrir *)
            nivelAlto := TRUE;
            tEspera   := T#3S;
            esperado  := TRUE;
        3:  (* Cae el nivel: debe cerrar de inmediato, sin retardo *)
            nivelAlto := FALSE;
            tEspera   := T#200MS;
            esperado  := FALSE;
        4:  (* Nuevo ciclo completo: comprueba el rearme del temporizador *)
            nivelAlto := TRUE;
            tEspera   := T#6S;
            esperado  := TRUE;
        5:  (* Cierre final *)
            nivelAlto := FALSE;
            tEspera   := T#200MS;
            esperado  := FALSE;
    END_CASE
END_IF

(* 2. Temporizador de asentamiento, con el tiempo propio del paso *)
tPaso(IN := NOT pulsoReset, PT := tEspera);
pulsoReset := FALSE;

(* 3. Llamada al bloque bajo prueba *)
fb(nivelAlto := nivelAlto);

(* 4. Evaluacion al vencer el asentamiento del paso *)
IF tPaso.Q AND NOT finalizado THEN
    IF fb.valvula = esperado THEN
        resultado[paso] := 1;
    ELSE
        resultado[paso] := 2;
    END_IF

    pulsoReset := TRUE;

    IF paso < ULTIMO_PASO THEN
        paso := paso + 1;
    ELSE
        finalizado := TRUE;
    END_IF
END_IF

(* 5. Veredicto global *)
IF finalizado AND veredicto = 0 THEN
    nPasan := 0;
    FOR i := 0 TO ULTIMO_PASO DO
        IF resultado[i] = 1 THEN
            nPasan := nPasan + 1;
        END_IF
    END_FOR

    IF nPasan = (ULTIMO_PASO + 1) THEN
        veredicto := 1;
    ELSE
        veredicto := 2;
    END_IF
END_IF

(* ---- PRG_Test_B3.st ---- *)
(*
    BANCO DE PRUEBA AUTOVERIFICABLE — Tarea B3 (contador de piezas por flanco)
    ---------------------------------------------------------------------------
    CORRIGE la version anterior, que tenia dos defectos fatales:

    1. El CASE asignaba sensorPieza := TRUE y una linea posterior lo invertia
       antes de llamar al bloque, de modo que el FB recibia siempre FALSE.
       No se generaba ningun flanco y el paso 4 reprobaba SIEMPRE, incluso a
       implementaciones correctas (falso negativo del 100%).

    2. La alternancia ocurria una vez por scan, por lo que el numero de flancos
       dependia del ciclo de la MainTask (2 flancos con 20 ms, 12 con 4 ms).
       El resultado era un accidente del entorno, no una medicion.

    SOLUCION: generador determinista de flancos con temporizador propio y
    contador explicito. Genera exactamente FLANCOS_EXTRA flancos ascendentes
    con independencia del ciclo de tarea. El temporizador de asentamiento del
    paso queda retenido mientras la generacion esta en curso, de modo que la
    evaluacion solo ocurre cuando ya se emitieron todos los flancos.

    3. (detectado por la validacion) Comprobar solo el estado final (cuenta=12,
       loteListo=TRUE) NO distingue un preset incorrecto: una implementacion que
       active el lote a las 10 piezas tambien llega a 12 con el lote activo. El
       umbral se verifica ahora en DOS LOTES: primero 10 flancos (cuenta=11, el
       lote debe seguir APAGADO) y despues 1 flanco mas (cuenta=12, lote ENCENDIDO).

    Cuentas esperadas: 1 (paso 1) + 10 (paso 4) + 1 (paso 5) = 12.
*)

PROGRAM PRG_Test_B3
VAR CONSTANT
    ULTIMO_PASO    : INT  := 6;
    FLANCOS_LOTE_A : INT  := 10;     (* 1 + 10 = 11 cuentas: el lote NO debe activarse *)
    FLANCOS_LOTE_B : INT  := 1;      (* 11 + 1 = 12 cuentas: el lote SI debe activarse *)
    T_PULSO        : TIME := T#20MS; (* semiperiodo del generador de flancos *)
END_VAR
VAR
    (* --- Bloque bajo prueba --- *)
    fb : FB_Contador;

    (* --- Entradas manipuladas por el banco --- *)
    sensorPieza : BOOL;
    btnReset    : BOOL;

    (* --- Control de la secuencia --- *)
    paso           : INT := 0;
    esperadoCuenta : INT;
    esperadoLote   : BOOL;
    tEspera        : TIME;
    tPaso          : TON;
    pulsoReset     : BOOL;
    finalizado     : BOOL;

    (* --- Generador determinista de flancos --- *)
    flancosPendientes : INT;
    pasoCargado       : INT := -1;   (* para cargar los flancos al entrar al paso *)
    tPulso            : TON;
    resetPulso        : BOOL;
    generando         : BOOL;

    (* --- Resultados --- *)
    resultado : ARRAY[0..6] OF INT;
    nPasan    : INT;
    veredicto : INT := 0;
    i         : INT;
END_VAR

(* 1. Definicion del paso en curso.
      En el paso 4 el CASE NO toca sensorPieza: lo gobierna el generador. *)
IF NOT finalizado THEN
    CASE paso OF
        0:  (* Reset inicial *)
            btnReset := TRUE;  sensorPieza := FALSE;
            tEspera := T#200MS; esperadoCuenta := 0; esperadoLote := FALSE;
        1:  (* Primer flanco ascendente *)
            btnReset := FALSE; sensorPieza := TRUE;
            tEspera := T#200MS; esperadoCuenta := 1; esperadoLote := FALSE;
        2:  (* Sensor sostenido en alto: NO debe seguir contando *)
            sensorPieza := TRUE;
            tEspera := T#500MS; esperadoCuenta := 1; esperadoLote := FALSE;
        3:  (* Vuelta a bajo para preparar la generacion *)
            sensorPieza := FALSE;
            tEspera := T#200MS; esperadoCuenta := 1; esperadoLote := FALSE;
        4:  (* 10 flancos -> 11 cuentas: el lote AUN NO debe activarse.
               Este paso es el que detecta un preset menor que 12. *)
            tEspera := T#200MS; esperadoCuenta := 11; esperadoLote := FALSE;
        5:  (* 1 flanco mas -> 12 cuentas: el lote SI debe activarse.
               Este paso detecta un preset mayor que 12. *)
            tEspera := T#200MS; esperadoCuenta := 12; esperadoLote := TRUE;
        6:  (* Reset final *)
            btnReset := TRUE;  sensorPieza := FALSE;
            tEspera := T#200MS; esperadoCuenta := 0; esperadoLote := FALSE;
    END_CASE
END_IF

(* 2. Carga del numero de flancos al entrar en cada paso generador *)
IF paso <> pasoCargado THEN
    CASE paso OF
        4: flancosPendientes := FLANCOS_LOTE_A;
        5: flancosPendientes := FLANCOS_LOTE_B;
    ELSE
        flancosPendientes := 0;
    END_CASE
    pasoCargado := paso;
END_IF

(* 3. Generador determinista de flancos (pasos 4 y 5) *)
generando := ((paso = 4) OR (paso = 5)) AND (flancosPendientes > 0);

IF generando THEN
    tPulso(IN := NOT resetPulso, PT := T_PULSO);
    resetPulso := FALSE;
    IF tPulso.Q THEN
        sensorPieza := NOT sensorPieza;
        IF sensorPieza THEN
            flancosPendientes := flancosPendientes - 1;   (* solo flancos ascendentes *)
        END_IF
        resetPulso := TRUE;
    END_IF
ELSE
    tPulso(IN := FALSE, PT := T_PULSO);
END_IF

(* 4. Asentamiento del paso, retenido mientras se generan flancos *)
tPaso(IN := NOT pulsoReset AND NOT generando, PT := tEspera);
pulsoReset := FALSE;

(* 5. Llamada al bloque bajo prueba *)
fb(sensorPieza := sensorPieza, btnReset := btnReset);

(* 6. Evaluacion al vencer el asentamiento *)
IF tPaso.Q AND NOT finalizado THEN
    IF (fb.cuenta = esperadoCuenta) AND (fb.loteListo = esperadoLote) THEN
        resultado[paso] := 1;
    ELSE
        resultado[paso] := 2;
    END_IF

    pulsoReset := TRUE;

    IF paso < ULTIMO_PASO THEN
        paso := paso + 1;
    ELSE
        finalizado := TRUE;
    END_IF
END_IF

(* 7. Veredicto global *)
IF finalizado AND veredicto = 0 THEN
    nPasan := 0;
    FOR i := 0 TO ULTIMO_PASO DO
        IF resultado[i] = 1 THEN
            nPasan := nPasan + 1;
        END_IF
    END_FOR

    IF nPasan = (ULTIMO_PASO + 1) THEN
        veredicto := 1;
    ELSE
        veredicto := 2;
    END_IF
END_IF

(* ---- PRG_Test_B4.st ---- *)
(*
    BANCO DE PRUEBA AUTOVERIFICABLE — Tarea B4 (inversion de giro)
    ---------------------------------------------------------------------------
    Propiedad critica (enmienda 4): "nunca fwd AND rev" se evalua en CADA scan
    y queda ENCLAVADA en 'violacionInterlock' hasta el final del banco, porque
    una violacion transitoria entre dos evaluaciones pasaria inadvertida. El
    veredicto final exige superar todos los pasos Y que la bandera este en
    FALSE. Se registra aparte porque una violacion de seguridad es
    cualitativamente distinta de un fallo funcional.

    USO: crear este PROGRAM junto al FUNCTION_BLOCK de la respuesta a evaluar y
    ejecutar en modo Simulacion. Al terminar, leer 'veredicto': 1 = supera,
    2 = falla.

    ---------------------------------------------------------------------------
    CORRECCION DEL 2026-09-09 (enmienda 9). Validado con validar_harness_B4.py.
    La version anterior daba veredicto 1, y sin levantar la bandera, a una
    implementacion con una CARRERA DE INTERLOCK: el enclavamiento cruzado se
    evaluaba contra el valor de la otra salida en el scan ANTERIOR. Con el
    motor ya girando se comporta bien, pero al pulsar las dos ordenes ESTANDO
    EN REPOSO ambas salidas se activan a la vez durante un scan.

    Causa: la secuencia solo pulsaba las dos ordenes con el motor ya girando en
    reversa (paso 6), situacion en la que la salida activa bloquea a la otra
    incluso con la comparacion retrasada. Nunca las pulsaba desde el reposo,
    que es justamente el caso en que la carrera se manifiesta.

    Es un fallo de COBERTURA, no del mecanismo: la enmienda 4 dejo el
    instrumento capaz de detectar la violacion transitoria, pero la secuencia
    no llegaba a provocarla. Una bandera enclavada solo puede atrapar lo que la
    secuencia produce.

    Correccion: se anaden dos pasos que pulsan ambas ordenes desde el reposo.
    El paso 8 no exige un sentido concreto —el enunciado no dice cual debe
    ganar si se piden los dos a la vez— sino unicamente que no coexistan.
*)

PROGRAM PRG_Test_B4
VAR CONSTANT
    ULTIMO_PASO    : INT  := 9;       (* 10 pasos: indices 0..9 *)
    T_ASENTAMIENTO : TIME := T#150MS;
END_VAR
VAR
    (* --- Bloque bajo prueba: sustituir por la respuesta a evaluar --- *)
    fb : FB_Giro;

    (* --- Entradas manipuladas por el banco --- *)
    btnFwd  : BOOL;
    btnRev  : BOOL;
    btnParo : BOOL;

    (* --- Control de la secuencia --- *)
    espFwd, espRev : BOOL;
    paso       : INT := 0;
    tPaso      : TON;
    pulsoReset : BOOL;
    finalizado : BOOL;

    (* --- Seguridad continua y enclavada (enmienda 4) --- *)
    violacionInterlock : BOOL;

    (* --- Resultados: 0 = pendiente, 1 = pasa, 2 = falla --- *)
    resultado : ARRAY[0..9] OF INT;
    nPasan    : INT;
    veredicto : INT := 0;
    i         : INT;
END_VAR

(* 1. Temporizador de asentamiento entre pasos *)
tPaso(IN := NOT pulsoReset, PT := T_ASENTAMIENTO);
pulsoReset := FALSE;

(* 2. Aplicacion de entradas y valores esperados. Solo se asigna lo que cada
      paso cambia: las demas entradas conservan su valor. *)
IF NOT finalizado THEN
    CASE paso OF
        0:  (* Reposo *)
            btnFwd := FALSE; btnRev := FALSE; btnParo := FALSE;
            espFwd := FALSE; espRev := FALSE;
        1:  (* Marcha adelante *)
            btnFwd := TRUE;
            espFwd := TRUE;  espRev := FALSE;
        2:  (* Se suelta la orden: debe mantenerse (enclavamiento) *)
            btnFwd := FALSE;
            espFwd := TRUE;  espRev := FALSE;
        3:  (* Reversa sin pasar por paro: prohibida *)
            btnRev := TRUE;
            espFwd := TRUE;  espRev := FALSE;
        4:  (* Paro *)
            btnRev := FALSE; btnParo := TRUE;
            espFwd := FALSE; espRev := FALSE;
        5:  (* Ahora si, marcha en reversa *)
            btnParo := FALSE; btnRev := TRUE;
            espFwd := FALSE; espRev := TRUE;
        6:  (* Ambas ordenes con el motor ya girando: la activa debe bloquear *)
            btnFwd := TRUE;
            espFwd := FALSE; espRev := TRUE;
        7:  (* Paro *)
            btnFwd := FALSE; btnRev := FALSE; btnParo := TRUE;
            espFwd := FALSE; espRev := FALSE;

        (* --- Ambas ordenes DESDE EL REPOSO (enmienda 9): es el unico caso en
               que una carrera de interlock se manifiesta --- *)
        8:  (* No se exige un sentido concreto, solo que no coexistan *)
            btnParo := FALSE; btnFwd := TRUE; btnRev := TRUE;
        9:  (* Paro final *)
            btnFwd := FALSE; btnRev := FALSE; btnParo := TRUE;
            espFwd := FALSE; espRev := FALSE;
    END_CASE
END_IF

(* 3. Llamada al bloque bajo prueba *)
fb(btnFwd := btnFwd, btnRev := btnRev, btnParo := btnParo);

(* 4. Seguridad: se evalua en CADA scan y queda enclavada (enmienda 4) *)
IF fb.fwd AND fb.rev THEN
    violacionInterlock := TRUE;
END_IF

(* 5. Evaluacion al vencer el asentamiento *)
IF tPaso.Q AND NOT finalizado THEN
    IF paso = 8 THEN
        (* El enunciado no fija cual de los dos sentidos debe ganar si se
           piden ambos a la vez, asi que el unico criterio es que no coexistan. *)
        IF NOT (fb.fwd AND fb.rev) THEN
            resultado[paso] := 1;
        ELSE
            resultado[paso] := 2;
        END_IF
    ELSE
        IF (fb.fwd = espFwd) AND (fb.rev = espRev) THEN
            resultado[paso] := 1;
        ELSE
            resultado[paso] := 2;
        END_IF
    END_IF

    pulsoReset := TRUE;

    IF paso < ULTIMO_PASO THEN
        paso := paso + 1;
    ELSE
        finalizado := TRUE;
    END_IF
END_IF

(* 6. Veredicto global: todos los pasos Y sin violacion de interlock *)
IF finalizado AND veredicto = 0 THEN
    nPasan := 0;
    FOR i := 0 TO ULTIMO_PASO DO
        IF resultado[i] = 1 THEN
            nPasan := nPasan + 1;
        END_IF
    END_FOR

    IF nPasan = (ULTIMO_PASO + 1) AND NOT violacionInterlock THEN
        veredicto := 1;
    ELSE
        veredicto := 2;
    END_IF
END_IF

(* ---- PRG_Test_B5.st ---- *)
(*
    BANCO DE PRUEBA AUTOVERIFICABLE — Tarea B5 (ventilador con retardo TOF)
    ---------------------------------------------------------------------------
    El ventilador acompana al quemador y sigue funcionando 30 s tras el paro.
    El punto delicado, declarado en ENMIENDAS_HARNESSES.md, es reactivar el
    quemador DURANTE el post-enfriamiento: la reactivacion debe REARMAR el
    temporizador, de modo que el siguiente post-enfriamiento vuelva a durar
    30 s completos.

    USO: crear este PROGRAM junto al FUNCTION_BLOCK de la respuesta a evaluar y
    ejecutar en modo Simulacion. Al terminar, leer 'veredicto': 1 = supera,
    2 = falla. 'resultado' indica el paso.

    ---------------------------------------------------------------------------
    CORRECCION DEL 2026-09-09 (enmienda 7). Validado con validar_harness_B5.py.
    La version anterior daba veredicto 1 a una implementacion que rearmaba el
    temporizador pero con un tiempo MENOR: el segundo post-enfriamiento duraba
    15 s en lugar de 30 s y pasaba como correcta en los tres ciclos de tarea.

    Causa: la secuencia reactivaba el quemador en el ultimo paso y terminaba
    ahi. Comprobaba que el temporizador se rearmaba, pero nunca que se rearmara
    a los 30 s completos, porque el segundo post-enfriamiento no se llegaba a
    recorrer. El paso final, ademas, no discriminaba nada: cualquier
    implementacion que superara el paso 1 lo superaba tambien.

    La propia enmienda de correccion de tiempos ya anticipaba esto al estimar
    B5 en ~70 s "porque la reactivacion durante el post-enfriamiento exige un
    segundo ciclo". La secuencia anterior duraba 41 s: el segundo ciclo que esa
    estimacion daba por hecho nunca se habia implementado.

    Correccion: tras la reactivacion se anaden dos pasos que recorren el
    segundo post-enfriamiento completo, con la misma pareja de comprobaciones
    que el primero (antes de los 30 s debe seguir encendido; pasados los 30 s
    debe estar apagado). La secuencia pasa a durar 71,2 s, acorde con la
    estimacion de la enmienda.
*)

PROGRAM PRG_Test_B5
VAR CONSTANT
    ULTIMO_PASO : INT := 8;          (* 9 pasos: indices 0..8 *)
END_VAR
VAR
    (* --- Bloque bajo prueba: sustituir por la respuesta a evaluar --- *)
    fb : FB_Ventilador;

    (* --- Entrada manipulada por el banco --- *)
    quemadorOn : BOOL;

    (* --- Control de la secuencia --- *)
    paso       : INT := 0;
    esperado   : BOOL;
    tEspera    : TIME;
    tPaso      : TON;
    pulsoReset : BOOL;
    finalizado : BOOL;

    (* --- Resultados: 0 = pendiente, 1 = pasa, 2 = falla --- *)
    resultado : ARRAY[0..8] OF INT;
    nPasan    : INT;
    veredicto : INT := 0;
    i         : INT;
END_VAR

(* 1. Definicion del paso en curso. Va antes del temporizador porque tEspera
      lo alimenta. *)
IF NOT finalizado THEN
    CASE paso OF
        0:  (* Reposo *)
            quemadorOn := FALSE; tEspera := T#200MS;  esperado := FALSE;
        1:  (* El ventilador acompana al quemador *)
            quemadorOn := TRUE;  tEspera := T#200MS;  esperado := TRUE;

        (* --- Primer post-enfriamiento --- *)
        2:  (* A los 29 s aun debe estar encendido *)
            quemadorOn := FALSE; tEspera := T#29S;    esperado := TRUE;
        3:  (* A los 30,2 s acumulados ya debe estar apagado *)
            quemadorOn := FALSE; tEspera := T#1200MS; esperado := FALSE;

        (* --- Reactivacion durante el post-enfriamiento --- *)
        4:  (* Se reenciende el quemador *)
            quemadorOn := TRUE;  tEspera := T#200MS;  esperado := TRUE;
        5:  (* Se apaga: arranca un post-enfriamiento que aun no vence *)
            quemadorOn := FALSE; tEspera := T#10S;    esperado := TRUE;
        6:  (* Se reenciende EN PLENO post-enfriamiento: debe rearmar *)
            quemadorOn := TRUE;  tEspera := T#200MS;  esperado := TRUE;

        (* --- Segundo post-enfriamiento COMPLETO (enmienda 7):
               no basta con que el temporizador se rearme, tiene que rearmarse
               a los 30 s completos --- *)
        7:  (* A los 29 s del nuevo paro aun debe estar encendido *)
            quemadorOn := FALSE; tEspera := T#29S;    esperado := TRUE;
        8:  (* A los 30,2 s del nuevo paro ya debe estar apagado *)
            quemadorOn := FALSE; tEspera := T#1200MS; esperado := FALSE;
    END_CASE
END_IF

(* 2. Temporizador de asentamiento del paso *)
tPaso(IN := NOT pulsoReset, PT := tEspera);
pulsoReset := FALSE;

(* 3. Llamada al bloque bajo prueba *)
fb(quemadorOn := quemadorOn);

(* 4. Evaluacion al vencer el asentamiento *)
IF tPaso.Q AND NOT finalizado THEN
    IF fb.ventilador = esperado THEN
        resultado[paso] := 1;
    ELSE
        resultado[paso] := 2;
    END_IF

    pulsoReset := TRUE;

    IF paso < ULTIMO_PASO THEN
        paso := paso + 1;
    ELSE
        finalizado := TRUE;
    END_IF
END_IF

(* 5. Veredicto global *)
IF finalizado AND veredicto = 0 THEN
    nPasan := 0;
    FOR i := 0 TO ULTIMO_PASO DO
        IF resultado[i] = 1 THEN
            nPasan := nPasan + 1;
        END_IF
    END_FOR

    IF nPasan = (ULTIMO_PASO + 1) THEN
        veredicto := 1;
    ELSE
        veredicto := 2;
    END_IF
END_IF

(* ---- PRG_Test_B6.st ---- *)
(*
    BANCO DE PRUEBA AUTOVERIFICABLE — Tarea B6 (baliza intermitente)
    ---------------------------------------------------------------------------
    Aplica la enmienda 1 de ENMIENDAS_HARNESSES.md: NO se muestrea la lampara,
    se MIDE la duracion de cada intervalo ON y OFF completo. Muestrear cada
    1,1 s no discrimina, porque una implementacion de 1,5 s / 1,5 s produce el
    mismo patron de alternancia que la correcta.

    El primer intervalo se descarta por parcial: depende de en que momento se
    activo la alarma. Se exige 1 s +/- 150 ms en al menos dos intervalos ON y
    dos OFF completos.

    Ciclo de MainTask: 4 a 10 ms (enmienda 3).

    USO: crear este PROGRAM junto al FUNCTION_BLOCK de la respuesta a evaluar y
    ejecutar en modo Simulacion. Al terminar, leer 'veredicto': 1 = supera,
    2 = falla. 'resultado' indica el paso.

    ---------------------------------------------------------------------------
    CORRECCION DEL 2026-09-09 (enmienda 6). Validado con validar_harness_B6.py.
    La version anterior daba veredicto 1 a una implementacion que SEGUIA
    PARPADEANDO despues de retirarse la alarma.

    Causa: el paso 2 esperaba 200 ms y comprobaba la lampara en un unico
    instante. Como la salida defectuosa es periodica, que se la sorprenda
    encendida o apagada depende de la fase en ese instante; en la simulacion
    caia sistematicamente en un tramo apagado y el defecto pasaba como bueno.
    Es exactamente el fallo de muestreo que la enmienda 1 corrigio para el
    paso 1, sin corregirse tambien en los pasos de reposo.

    Correccion, con la misma logica de la enmienda 4: la condicion se evalua en
    CADA scan y queda ENCLAVADA, y la ventana del paso 2 pasa de 200 ms a
    2,5 s, mas de dos periodos nominales completos. Asi cualquier parpadeo
    indebido con semiperiodo por debajo de ~2,5 s queda registrado.

    Se unifica ademas la medida de intervalos con el metodo adoptado en la
    enmienda 5 para I4: diferencia de dos lecturas de un cronometro libre, en
    lugar de reiniciar un temporizador con un ciclo de retraso. Con la
    tolerancia de +/- 150 ms el sesgo anterior no llegaba a ser un defecto
    (medía ~980 ms en vez de 1000 ms con ciclo de 20 ms), pero no hay razon
    para conservar un sesgo conocido.
*)

PROGRAM PRG_Test_B6
VAR CONSTANT
    ULTIMO_PASO : INT  := 2;
    T_NOMINAL   : TIME := T#1S;
    TOL_MIN     : TIME := T#850MS;    (* 1 s - 150 ms *)
    TOL_MAX     : TIME := T#1150MS;   (* 1 s + 150 ms *)
    T_REPOSO    : TIME := T#2500MS;   (* > 2 periodos nominales (enmienda 6) *)
    T_CRONO     : TIME := T#100S;     (* cronometro libre: nunca se reinicia *)
END_VAR
VAR
    (* --- Bloque bajo prueba: sustituir por la respuesta a evaluar --- *)
    fb : FB_Baliza;

    (* --- Entrada manipulada por el banco --- *)
    alarma : BOOL;

    (* --- Control de la secuencia --- *)
    paso       : INT := 0;
    tEspera    : TIME;
    tPaso      : TON;
    pulsoReset : BOOL;
    finalizado : BOOL;

    (* --- Medida de intervalos (enmienda 1) --- *)
    tCrono       : TON;
    prev         : BOOL;
    primer       : BOOL;              (* el primer intervalo es parcial *)
    etFlanco     : TIME;
    duracion     : TIME;
    error        : BOOL;              (* algun intervalo fuera de tolerancia *)
    nOn, nOff    : INT;

    (* --- Vigilancia de reposo, continua y enclavada (enmienda 6) --- *)
    lamparaEnPaso0 : BOOL;
    lamparaEnPaso2 : BOOL;

    (* --- Resultados: 0 = pendiente, 1 = pasa, 2 = falla --- *)
    resultado : ARRAY[0..2] OF INT;
    nPasan    : INT;
    veredicto : INT := 0;
    i         : INT;
END_VAR

(* 1. Definicion del paso en curso *)
IF NOT finalizado THEN
    CASE paso OF
        0:  (* Reposo inicial: sin alarma, la lampara debe estar apagada *)
            alarma  := FALSE;
            tEspera := T#200MS;
        1:  (* Alarma activa: ventana de observacion del parpadeo *)
            alarma  := TRUE;
            tEspera := T#7S;
        2:  (* Alarma retirada: debe apagarse y PERMANECER apagada *)
            alarma  := FALSE;
            tEspera := T_REPOSO;
    END_CASE
END_IF

(* 2. Temporizadores del banco *)
tPaso(IN := NOT pulsoReset, PT := tEspera);
tCrono(IN := TRUE, PT := T_CRONO);
pulsoReset := FALSE;

(* 3. Llamada al bloque bajo prueba *)
fb(alarma := alarma);

(* 4. Medida de intervalos completos durante el paso 1 (enmienda 1).
      La duracion se obtiene por diferencia de dos lecturas del cronometro
      libre, no reiniciando un temporizador (enmienda 5). *)
IF paso = 1 THEN
    IF (fb.lampara AND NOT prev) OR ((NOT fb.lampara) AND prev) THEN
        IF primer THEN
            duracion := tCrono.ET - etFlanco;
            IF NOT fb.lampara THEN
                nOn := nOn + 1;        (* se acaba de cerrar un intervalo ON *)
            ELSE
                nOff := nOff + 1;      (* se acaba de cerrar un intervalo OFF *)
            END_IF
            IF duracion < TOL_MIN OR duracion > TOL_MAX THEN
                error := TRUE;
            END_IF
        ELSE
            primer := TRUE;            (* se descarta el intervalo parcial *)
        END_IF
        etFlanco := tCrono.ET;
    END_IF
END_IF

(* 5. Vigilancia de reposo: se evalua en CADA scan y queda enclavada
      (enmienda 6). Un unico muestreo al final del paso no sirve porque la
      salida defectuosa es periodica. *)
IF paso = 0 AND fb.lampara THEN
    lamparaEnPaso0 := TRUE;
END_IF
IF paso = 2 AND fb.lampara THEN
    lamparaEnPaso2 := TRUE;
END_IF

prev := fb.lampara;

(* 6. Evaluacion al vencer el asentamiento del paso *)
IF tPaso.Q AND NOT finalizado THEN
    IF    (paso = 0 AND NOT fb.lampara AND NOT lamparaEnPaso0)
       OR (paso = 1 AND nOn >= 2 AND nOff >= 2 AND NOT error)
       OR (paso = 2 AND NOT fb.lampara AND NOT lamparaEnPaso2)
    THEN
        resultado[paso] := 1;
    ELSE
        resultado[paso] := 2;
    END_IF

    pulsoReset := TRUE;

    IF paso < ULTIMO_PASO THEN
        paso := paso + 1;
    ELSE
        finalizado := TRUE;
    END_IF
END_IF

(* 7. Veredicto global *)
IF finalizado AND veredicto = 0 THEN
    nPasan := 0;
    FOR i := 0 TO ULTIMO_PASO DO
        IF resultado[i] = 1 THEN
            nPasan := nPasan + 1;
        END_IF
    END_FOR

    IF nPasan = (ULTIMO_PASO + 1) THEN
        veredicto := 1;
    ELSE
        veredicto := 2;
    END_IF
END_IF

(* ---- PRG_Test_B7_FB.st ---- *)
(*
    BANCO DE PRUEBA AUTOVERIFICABLE - Tarea B7 (SelBomba, POU a eleccion)
    VARIANTE: FUNCTION_BLOCK  (generada por generar_harness_B7.py; no editar a mano)
    ---------------------------------------------------------------------------
    Validado en codesys/validar_harness_B7.py: 9 implementaciones (3 correctas,
    una por tipo de POU, y 6 defectuosas), ciclos de 4, 10 y 20 ms.
    Las tres variantes comparten secuencia y evaluacion; solo cambia la llamada.

    Paso (modoAuto, btnManual, nivelBajo) -> bomba
      0 (F,F,F) F   1 (F,T,F) T   2 (F,F,F) F   3 (F,F,T) F   4 (T,F,T) T
      5 (T,F,F) F   6 (T,T,F) F   7 (T,T,T) T   8 (F,T,T) T   9 (F,F,T) F
    Cada paso de TRUE a FALSE delata memoria entre ciclos (el enunciado la prohibe).
*)
PROGRAM PRG_Test_B7
VAR CONSTANT
    ULTIMO_PASO : INT  := 9;
    T_PASO      : TIME := T#100MS;
END_VAR
VAR
    fb : SelBomba;           (* instancia del FB bajo prueba *)
    modoAuto   : BOOL;
    btnManual  : BOOL;
    nivelBajo  : BOOL;
    bomba      : BOOL;       (* salida leida del POU bajo prueba *)
    esperado   : BOOL;

    paso       : INT := 0;
    tPaso      : TON;
    pulsoReset : BOOL;
    finalizado : BOOL;

    resultado : ARRAY[0..9] OF INT;
    nPasan    : INT;
    veredicto : INT := 0;
    i         : INT;
END_VAR

(* 1. Entradas y valor esperado del paso *)
IF NOT finalizado THEN
    CASE paso OF
        0: modoAuto := FALSE; btnManual := FALSE; nivelBajo := FALSE; esperado := FALSE;
        1: modoAuto := FALSE; btnManual := TRUE;  nivelBajo := FALSE; esperado := TRUE;
        2: modoAuto := FALSE; btnManual := FALSE; nivelBajo := FALSE; esperado := FALSE;
        3: modoAuto := FALSE; btnManual := FALSE; nivelBajo := TRUE;  esperado := FALSE;
        4: modoAuto := TRUE;  btnManual := FALSE; nivelBajo := TRUE;  esperado := TRUE;
        5: modoAuto := TRUE;  btnManual := FALSE; nivelBajo := FALSE; esperado := FALSE;
        6: modoAuto := TRUE;  btnManual := TRUE;  nivelBajo := FALSE; esperado := FALSE;
        7: modoAuto := TRUE;  btnManual := TRUE;  nivelBajo := TRUE;  esperado := TRUE;
        8: modoAuto := FALSE; btnManual := TRUE;  nivelBajo := TRUE;  esperado := TRUE;
        9: modoAuto := FALSE; btnManual := FALSE; nivelBajo := TRUE;  esperado := FALSE;
    END_CASE
END_IF

(* 2. Asentamiento del paso *)
tPaso(IN := NOT pulsoReset, PT := T_PASO);
pulsoReset := FALSE;

(* 3. Llamada al POU bajo prueba (FUNCTION_BLOCK) *)
fb(modoAuto := modoAuto, btnManual := btnManual, nivelBajo := nivelBajo);
bomba := fb.bomba;

(* 4. Evaluacion *)
IF tPaso.Q AND NOT finalizado THEN
    IF bomba = esperado THEN
        resultado[paso] := 1;
    ELSE
        resultado[paso] := 2;
    END_IF
    pulsoReset := TRUE;
    IF paso < ULTIMO_PASO THEN
        paso := paso + 1;
    ELSE
        finalizado := TRUE;
    END_IF
END_IF

(* 5. Veredicto global *)
IF finalizado AND veredicto = 0 THEN
    nPasan := 0;
    FOR i := 0 TO ULTIMO_PASO DO
        IF resultado[i] = 1 THEN
            nPasan := nPasan + 1;
        END_IF
    END_FOR
    IF nPasan = (ULTIMO_PASO + 1) THEN
        veredicto := 1;
    ELSE
        veredicto := 2;
    END_IF
END_IF

(* ---- PRG_Test_B7_FUN.st ---- *)
(*
    BANCO DE PRUEBA AUTOVERIFICABLE - Tarea B7 (SelBomba, POU a eleccion)
    VARIANTE: FUNCTION  (generada por generar_harness_B7.py; no editar a mano)
    ---------------------------------------------------------------------------
    Validado en codesys/validar_harness_B7.py: 9 implementaciones (3 correctas,
    una por tipo de POU, y 6 defectuosas), ciclos de 4, 10 y 20 ms.
    Las tres variantes comparten secuencia y evaluacion; solo cambia la llamada.

    Paso (modoAuto, btnManual, nivelBajo) -> bomba
      0 (F,F,F) F   1 (F,T,F) T   2 (F,F,F) F   3 (F,F,T) F   4 (T,F,T) T
      5 (T,F,F) F   6 (T,T,F) F   7 (T,T,T) T   8 (F,T,T) T   9 (F,F,T) F
    Cada paso de TRUE a FALSE delata memoria entre ciclos (el enunciado la prohibe).
*)
PROGRAM PRG_Test_B7
VAR CONSTANT
    ULTIMO_PASO : INT  := 9;
    T_PASO      : TIME := T#100MS;
END_VAR
VAR
    (* sin instancia: SelBomba es una FUNCTION *)
    modoAuto   : BOOL;
    btnManual  : BOOL;
    nivelBajo  : BOOL;
    bomba      : BOOL;       (* salida leida del POU bajo prueba *)
    esperado   : BOOL;

    paso       : INT := 0;
    tPaso      : TON;
    pulsoReset : BOOL;
    finalizado : BOOL;

    resultado : ARRAY[0..9] OF INT;
    nPasan    : INT;
    veredicto : INT := 0;
    i         : INT;
END_VAR

(* 1. Entradas y valor esperado del paso *)
IF NOT finalizado THEN
    CASE paso OF
        0: modoAuto := FALSE; btnManual := FALSE; nivelBajo := FALSE; esperado := FALSE;
        1: modoAuto := FALSE; btnManual := TRUE;  nivelBajo := FALSE; esperado := TRUE;
        2: modoAuto := FALSE; btnManual := FALSE; nivelBajo := FALSE; esperado := FALSE;
        3: modoAuto := FALSE; btnManual := FALSE; nivelBajo := TRUE;  esperado := FALSE;
        4: modoAuto := TRUE;  btnManual := FALSE; nivelBajo := TRUE;  esperado := TRUE;
        5: modoAuto := TRUE;  btnManual := FALSE; nivelBajo := FALSE; esperado := FALSE;
        6: modoAuto := TRUE;  btnManual := TRUE;  nivelBajo := FALSE; esperado := FALSE;
        7: modoAuto := TRUE;  btnManual := TRUE;  nivelBajo := TRUE;  esperado := TRUE;
        8: modoAuto := FALSE; btnManual := TRUE;  nivelBajo := TRUE;  esperado := TRUE;
        9: modoAuto := FALSE; btnManual := FALSE; nivelBajo := TRUE;  esperado := FALSE;
    END_CASE
END_IF

(* 2. Asentamiento del paso *)
tPaso(IN := NOT pulsoReset, PT := T_PASO);
pulsoReset := FALSE;

(* 3. Llamada al POU bajo prueba (FUNCTION) *)
bomba := SelBomba(modoAuto := modoAuto, btnManual := btnManual, nivelBajo := nivelBajo);

(* 4. Evaluacion *)
IF tPaso.Q AND NOT finalizado THEN
    IF bomba = esperado THEN
        resultado[paso] := 1;
    ELSE
        resultado[paso] := 2;
    END_IF
    pulsoReset := TRUE;
    IF paso < ULTIMO_PASO THEN
        paso := paso + 1;
    ELSE
        finalizado := TRUE;
    END_IF
END_IF

(* 5. Veredicto global *)
IF finalizado AND veredicto = 0 THEN
    nPasan := 0;
    FOR i := 0 TO ULTIMO_PASO DO
        IF resultado[i] = 1 THEN
            nPasan := nPasan + 1;
        END_IF
    END_FOR
    IF nPasan = (ULTIMO_PASO + 1) THEN
        veredicto := 1;
    ELSE
        veredicto := 2;
    END_IF
END_IF

(* ---- PRG_Test_B7_PRG.st ---- *)
(*
    BANCO DE PRUEBA AUTOVERIFICABLE - Tarea B7 (SelBomba, POU a eleccion)
    VARIANTE: PROGRAM  (generada por generar_harness_B7.py; no editar a mano)
    ---------------------------------------------------------------------------
    Validado en codesys/validar_harness_B7.py: 9 implementaciones (3 correctas,
    una por tipo de POU, y 6 defectuosas), ciclos de 4, 10 y 20 ms.
    Las tres variantes comparten secuencia y evaluacion; solo cambia la llamada.

    Paso (modoAuto, btnManual, nivelBajo) -> bomba
      0 (F,F,F) F   1 (F,T,F) T   2 (F,F,F) F   3 (F,F,T) F   4 (T,F,T) T
      5 (T,F,F) F   6 (T,T,F) F   7 (T,T,T) T   8 (F,T,T) T   9 (F,F,T) F
    Cada paso de TRUE a FALSE delata memoria entre ciclos (el enunciado la prohibe).
*)
PROGRAM PRG_Test_B7
VAR CONSTANT
    ULTIMO_PASO : INT  := 9;
    T_PASO      : TIME := T#100MS;
END_VAR
VAR
    (* sin instancia: SelBomba es un PROGRAM, se llama por su nombre *)
    modoAuto   : BOOL;
    btnManual  : BOOL;
    nivelBajo  : BOOL;
    bomba      : BOOL;       (* salida leida del POU bajo prueba *)
    esperado   : BOOL;

    paso       : INT := 0;
    tPaso      : TON;
    pulsoReset : BOOL;
    finalizado : BOOL;

    resultado : ARRAY[0..9] OF INT;
    nPasan    : INT;
    veredicto : INT := 0;
    i         : INT;
END_VAR

(* 1. Entradas y valor esperado del paso *)
IF NOT finalizado THEN
    CASE paso OF
        0: modoAuto := FALSE; btnManual := FALSE; nivelBajo := FALSE; esperado := FALSE;
        1: modoAuto := FALSE; btnManual := TRUE;  nivelBajo := FALSE; esperado := TRUE;
        2: modoAuto := FALSE; btnManual := FALSE; nivelBajo := FALSE; esperado := FALSE;
        3: modoAuto := FALSE; btnManual := FALSE; nivelBajo := TRUE;  esperado := FALSE;
        4: modoAuto := TRUE;  btnManual := FALSE; nivelBajo := TRUE;  esperado := TRUE;
        5: modoAuto := TRUE;  btnManual := FALSE; nivelBajo := FALSE; esperado := FALSE;
        6: modoAuto := TRUE;  btnManual := TRUE;  nivelBajo := FALSE; esperado := FALSE;
        7: modoAuto := TRUE;  btnManual := TRUE;  nivelBajo := TRUE;  esperado := TRUE;
        8: modoAuto := FALSE; btnManual := TRUE;  nivelBajo := TRUE;  esperado := TRUE;
        9: modoAuto := FALSE; btnManual := FALSE; nivelBajo := TRUE;  esperado := FALSE;
    END_CASE
END_IF

(* 2. Asentamiento del paso *)
tPaso(IN := NOT pulsoReset, PT := T_PASO);
pulsoReset := FALSE;

(* 3. Llamada al POU bajo prueba (PROGRAM) *)
SelBomba(modoAuto := modoAuto, btnManual := btnManual, nivelBajo := nivelBajo);
bomba := SelBomba.bomba;

(* 4. Evaluacion *)
IF tPaso.Q AND NOT finalizado THEN
    IF bomba = esperado THEN
        resultado[paso] := 1;
    ELSE
        resultado[paso] := 2;
    END_IF
    pulsoReset := TRUE;
    IF paso < ULTIMO_PASO THEN
        paso := paso + 1;
    ELSE
        finalizado := TRUE;
    END_IF
END_IF

(* 5. Veredicto global *)
IF finalizado AND veredicto = 0 THEN
    nPasan := 0;
    FOR i := 0 TO ULTIMO_PASO DO
        IF resultado[i] = 1 THEN
            nPasan := nPasan + 1;
        END_IF
    END_FOR
    IF nPasan = (ULTIMO_PASO + 1) THEN
        veredicto := 1;
    ELSE
        veredicto := 2;
    END_IF
END_IF

(* ---- PRG_Test_B8.st ---- *)
(*
    BANCO DE PRUEBA AUTOVERIFICABLE - Tarea B8 (FB_Puerta: aperturas por flanco)
    ---------------------------------------------------------------------------
    Validado por simulacion en codesys/validar_harness_B8.py (traduccion fiel):
    9 implementaciones (1 correcta, 8 defectuosas), ciclos de 4, 10 y 20 ms.

    Pasos (cuentas acumuladas):
      0 reset, puerta cerrada ............................ n=0  aviso=F
      1 se suelta reset y se abre la puerta (1 flanco) ... n=1  aviso=F
      2 puerta sostenida abierta 500 ms .................. n=1  aviso=F
      3 puerta cerrada ................................... n=1  aviso=F
      4 3 flancos generados .............................. n=4  aviso=F  (umbral 4)
      5 1 flanco ......................................... n=5  aviso=T  (umbral '>5')
      6 1 flanco ......................................... n=6  aviso=T  ('=5', saturacion)
      7 reset, puerta cerrada ............................ n=0  aviso=F  (reset incompleto)
      8 se suelta reset, 1 flanco ........................ n=1  aviso=F  (bloqueo tras reset)
    Las transiciones de reset se hacen con la puerta cerrada: el enunciado no
    define que pasa con un flanco durante el reset, asi que no se prueba.

    Generador determinista de flancos (patron de B3): el numero de flancos no
    depende del ciclo de la MainTask; el asentamiento del paso queda retenido
    mientras se generan.
*)
PROGRAM PRG_Test_B8
VAR CONSTANT
    ULTIMO_PASO : INT  := 8;
    T_PULSO     : TIME := T#20MS;
END_VAR
VAR
    fb : FB_Puerta;                 (* bloque bajo prueba *)

    puertaAbierta : BOOL;
    reset         : BOOL;

    paso        : INT := 0;
    esperadoN   : INT;
    esperadoAv  : BOOL;
    tEspera     : TIME;
    tPaso       : TON;
    pulsoReset  : BOOL;
    finalizado  : BOOL;

    flancosPendientes : INT;
    pasoCargado       : INT := -1;
    tPulso            : TON;
    resetPulso        : BOOL;
    generando         : BOOL;

    resultado : ARRAY[0..8] OF INT;
    nPasan    : INT;
    veredicto : INT := 0;
    i         : INT;
END_VAR

(* 1. Definicion del paso. En los pasos 4, 5, 6 y 8 la puerta la gobierna el generador. *)
IF NOT finalizado THEN
    CASE paso OF
        0: reset := TRUE;  puertaAbierta := FALSE; tEspera := T#200MS; esperadoN := 0; esperadoAv := FALSE;
        1: reset := FALSE; puertaAbierta := TRUE;  tEspera := T#200MS; esperadoN := 1; esperadoAv := FALSE;
        2: puertaAbierta := TRUE;                  tEspera := T#500MS; esperadoN := 1; esperadoAv := FALSE;
        3: puertaAbierta := FALSE;                 tEspera := T#200MS; esperadoN := 1; esperadoAv := FALSE;
        4:                                         tEspera := T#200MS; esperadoN := 4; esperadoAv := FALSE;
        5:                                         tEspera := T#200MS; esperadoN := 5; esperadoAv := TRUE;
        6:                                         tEspera := T#200MS; esperadoN := 6; esperadoAv := TRUE;
        7: reset := TRUE;  puertaAbierta := FALSE; tEspera := T#200MS; esperadoN := 0; esperadoAv := FALSE;
        8: reset := FALSE;                         tEspera := T#200MS; esperadoN := 1; esperadoAv := FALSE;
    END_CASE
END_IF

(* 2. Carga del numero de flancos al entrar en cada paso *)
IF paso <> pasoCargado THEN
    CASE paso OF
        4: flancosPendientes := 3;
        5, 6, 8: flancosPendientes := 1;
    ELSE
        flancosPendientes := 0;
    END_CASE
    pasoCargado := paso;
END_IF

(* 3. Generador determinista de flancos *)
generando := flancosPendientes > 0;
IF generando THEN
    tPulso(IN := NOT resetPulso, PT := T_PULSO);
    resetPulso := FALSE;
    IF tPulso.Q THEN
        puertaAbierta := NOT puertaAbierta;
        IF puertaAbierta THEN
            flancosPendientes := flancosPendientes - 1;   (* solo flancos ascendentes *)
        END_IF
        resetPulso := TRUE;
    END_IF
ELSE
    tPulso(IN := FALSE, PT := T_PULSO);
END_IF

(* 4. Asentamiento, retenido mientras se generan flancos *)
tPaso(IN := NOT pulsoReset AND NOT generando, PT := tEspera);
pulsoReset := FALSE;

(* 5. Bloque bajo prueba *)
fb(puertaAbierta := puertaAbierta, reset := reset);

(* 6. Evaluacion *)
IF tPaso.Q AND NOT finalizado THEN
    IF (fb.nAperturas = esperadoN) AND (fb.aviso = esperadoAv) THEN
        resultado[paso] := 1;
    ELSE
        resultado[paso] := 2;
    END_IF
    pulsoReset := TRUE;
    IF paso < ULTIMO_PASO THEN
        paso := paso + 1;
    ELSE
        finalizado := TRUE;
    END_IF
END_IF

(* 7. Veredicto global *)
IF finalizado AND veredicto = 0 THEN
    nPasan := 0;
    FOR i := 0 TO ULTIMO_PASO DO
        IF resultado[i] = 1 THEN
            nPasan := nPasan + 1;
        END_IF
    END_FOR
    IF nPasan = (ULTIMO_PASO + 1) THEN
        veredicto := 1;
    ELSE
        veredicto := 2;
    END_IF
END_IF

(* ---- PRG_Test_C3.st ---- *)
(*
    BANCO DE PRUEBA AUTOVERIFICABLE - Tarea C3 (conversion Ladder -> ST, PRG_Conversion)
    ---------------------------------------------------------------------------
    Validado en codesys/validar_harness_C3.py: 7 implementaciones (1 correcta y
    6 defectuosas), ciclos de 4, 10 y 20 ms. Tabla de pasos generada desde el
    validador. Una respuesta con las E/S en VAR local no compila con este banco
    (CODESYS no admite escribir desde fuera una VAR local de un PROGRAM): se
    clasifica como INTERFAZ NO CONFORME, igual que los FB con E/S en VAR.
    El POU bajo prueba es un PROGRAM: se escriben sus entradas y se leen sus
    salidas por nombre, y se llama una vez por scan desde este banco.

    Paso (btnMarcha, btnParo) duracion -> (motor, lampara)
  0 (F,F) 0.2 s -> (F,F)
  1 (T,F) 0.2 s -> (T,F)   arranque; la lampara aun no
  2 (F,F) 5.0 s -> (T,F)   enclavamiento; lampara vigilada en FALSE todo el paso
  3 (F,F) 5.5 s -> (T,T)   ~10.7 s con motor: lampara encendida
  4 (F,T) 0.2 s -> (F,F)   paro: motor y lampara (T1 se reinicia)
  5 (F,F) 0.2 s -> (F,F)
  6 (T,T) 0.2 s -> (F,F)   marcha y paro a la vez: gana el NC en serie; vigilado
  7 (T,F) 0.2 s -> (T,F)
  8 (F,F) 9.0 s -> (T,F)   T1 empezo de cero en el paso 7: lampara vigilada en FALSE
  9 (F,F) 1.5 s -> (T,T)
 10 (F,T) 0.2 s -> (F,F)
VIGILANCIA CONTINUA (enmienda 4): en los pasos 0, 2, 5, 6 y 8 la lampara no puede
valer TRUE ni un scan; en los pasos 0, 5 y 6 tampoco el motor.
*)
PROGRAM PRG_Test_C3
VAR CONSTANT
    ULTIMO_PASO : INT := 10;
END_VAR
VAR
    bM, bP             : BOOL;     (* btnMarcha, btnParo aplicados *)
    eMotor, eLampara   : BOOL;     (* esperados *)

    paso       : INT := 0;
    tEspera    : TIME;
    tPaso      : TON;
    pulsoReset : BOOL;
    finalizado : BOOL;
    vigLampara : BOOL;
    vigMotor   : BOOL;
    violacion  : BOOL;

    resultado : ARRAY[0..10] OF INT;
    nPasan    : INT;
    veredicto : INT := 0;
    i         : INT;
END_VAR

(* 1. Entradas, duracion y salidas esperadas del paso *)
IF NOT finalizado THEN
    CASE paso OF
        0: bM := FALSE; bP := FALSE; tEspera := T#200MS; eMotor := FALSE; eLampara := FALSE;
        1: bM := TRUE; bP := FALSE; tEspera := T#200MS; eMotor := TRUE; eLampara := FALSE;
        2: bM := FALSE; bP := FALSE; tEspera := T#5000MS; eMotor := TRUE; eLampara := FALSE;
        3: bM := FALSE; bP := FALSE; tEspera := T#5500MS; eMotor := TRUE; eLampara := TRUE;
        4: bM := FALSE; bP := TRUE; tEspera := T#200MS; eMotor := FALSE; eLampara := FALSE;
        5: bM := FALSE; bP := FALSE; tEspera := T#200MS; eMotor := FALSE; eLampara := FALSE;
        6: bM := TRUE; bP := TRUE; tEspera := T#200MS; eMotor := FALSE; eLampara := FALSE;
        7: bM := TRUE; bP := FALSE; tEspera := T#200MS; eMotor := TRUE; eLampara := FALSE;
        8: bM := FALSE; bP := FALSE; tEspera := T#9000MS; eMotor := TRUE; eLampara := FALSE;
        9: bM := FALSE; bP := FALSE; tEspera := T#1500MS; eMotor := TRUE; eLampara := TRUE;
        10: bM := FALSE; bP := TRUE; tEspera := T#200MS; eMotor := FALSE; eLampara := FALSE;
    END_CASE
END_IF

(* 2. Asentamiento del paso *)
tPaso(IN := NOT pulsoReset, PT := tEspera);
pulsoReset := FALSE;

(* 3. PROGRAM bajo prueba *)
PRG_Conversion.btnMarcha := bM;
PRG_Conversion.btnParo := bP;
PRG_Conversion();

(* 4. Vigilancia continua *)
CASE paso OF
    0, 2, 5, 6, 8: vigLampara := TRUE;
ELSE
    vigLampara := FALSE;
END_CASE
CASE paso OF
    0, 5, 6: vigMotor := TRUE;
ELSE
    vigMotor := FALSE;
END_CASE
IF NOT finalizado AND ((vigLampara AND PRG_Conversion.lampara) OR (vigMotor AND PRG_Conversion.motor)) THEN
    violacion := TRUE;
END_IF

(* 5. Evaluacion *)
IF tPaso.Q AND NOT finalizado THEN
    IF (PRG_Conversion.motor = eMotor) AND (PRG_Conversion.lampara = eLampara) AND NOT violacion THEN
        resultado[paso] := 1;
    ELSE
        resultado[paso] := 2;
    END_IF
    violacion := FALSE;
    pulsoReset := TRUE;
    IF paso < ULTIMO_PASO THEN
        paso := paso + 1;
    ELSE
        finalizado := TRUE;
    END_IF
END_IF

(* 6. Veredicto global *)
IF finalizado AND veredicto = 0 THEN
    nPasan := 0;
    FOR i := 0 TO ULTIMO_PASO DO
        IF resultado[i] = 1 THEN
            nPasan := nPasan + 1;
        END_IF
    END_FOR
    IF nPasan = (ULTIMO_PASO + 1) THEN
        veredicto := 1;
    ELSE
        veredicto := 2;
    END_IF
END_IF

(* ---- PRG_Test_I1.st ---- *)
(*
    BANCO DE PRUEBA AUTOVERIFICABLE — Tarea I1 (semaforo con secuencia temporizada)
    ---------------------------------------------------------------------------
    Verde 20 s, amarillo 4 s, rojo 15 s, ciclico mientras 'habilitado'. Al
    deshabilitar, amarillo intermitente de 1 s / 1 s con las demas luces
    apagadas. Al rehabilitar, la secuencia REINICIA EN VERDE.

    El modo intermitente se verifica midiendo la duracion de los intervalos
    completos, no muestreando (enmienda 1). La condicion "las demas luces
    apagadas" se vigila en cada scan y queda enclavada (enmienda 6).

    Ciclo de MainTask: 4 a 10 ms (enmienda 3).

    USO: crear este PROGRAM junto al FUNCTION_BLOCK de la respuesta a evaluar y
    ejecutar en modo Simulacion. Al terminar, leer 'veredicto': 1 = supera,
    2 = falla. 'resultado' indica el paso.

    ---------------------------------------------------------------------------
    CORRECCION DEL 2026-09-09 (enmienda 8). Validado con validar_harness_I1.py.
    La version anterior daba veredicto 1 a dos implementaciones defectuosas:

    FALLO 1 — "las demas luces apagadas" se comprobaba en un unico instante al
    final del paso intermitente. Una implementacion que resuelve el
    intermitente alternando AMARILLO y ROJO (error plausible: parpadear entre
    el amarillo y la ultima luz activa) deja el rojo en antifase con el
    amarillo, de modo que en el instante muestreado las demas estan apagadas.
    Verificado: con el parpadeo arrancando en amarillo encendido, el defecto
    obtiene veredicto 1 en los tres ciclos de tarea; con la fase contraria solo
    se detecta de rebote en el paso 0, es decir por suerte de fase y no por
    merito del banco. Es el mismo error de muestreo de la enmienda 6.

    FALLO 2 — el reinicio en verde no se estaba probando. La secuencia
    deshabilitaba el semaforo mientras estaba EN VERDE, asi que al rehabilitar
    una implementacion que reinicia y una que continua donde se quedo muestran
    exactamente lo mismo. Verificado: el defecto "no reinicia" obtenia
    veredicto 1 en los tres ciclos. Para probarlo hay que interrumpir en una
    fase que NO sea verde.

    Correcciones: la vigilancia de V y R en los pasos deshabilitados pasa a ser
    continua y enclavada; y la secuencia recorre un segundo ciclo hasta el ROJO
    antes de deshabilitar, de modo que el reinicio en verde sea observable. La
    medida de intervalos se unifica con el metodo de la enmienda 5 (diferencia
    de dos lecturas de un cronometro libre). La secuencia pasa de 46,6 s a
    70,6 s, dentro de la estimacion de ~90 s de la correccion de tiempos.
*)

PROGRAM PRG_Test_I1
VAR CONSTANT
    ULTIMO_PASO : INT  := 8;          (* 9 pasos: indices 0..8 *)
    TOL_MIN     : TIME := T#850MS;    (* 1 s - 150 ms *)
    TOL_MAX     : TIME := T#1150MS;   (* 1 s + 150 ms *)
    T_CRONO     : TIME := T#100S;
END_VAR
VAR
    (* --- Bloque bajo prueba: sustituir por la respuesta a evaluar --- *)
    fb : FB_Semaforo;

    (* --- Entrada manipulada por el banco --- *)
    habilitado : BOOL;

    (* --- Control de la secuencia --- *)
    paso       : INT := 0;
    tEspera    : TIME;
    espV, espA, espR : BOOL;
    tPaso      : TON;
    pulsoReset : BOOL;
    finalizado : BOOL;

    (* --- Medida del intermitente (enmiendas 1 y 5) --- *)
    tCrono   : TON;
    prevA    : BOOL;
    primer   : BOOL;
    etFlanco : TIME;
    duracion : TIME;
    error    : BOOL;
    nOn, nOff : INT;

    (* --- Vigilancia continua y enclavada de las demas luces (enmienda 6) --- *)
    otraLuzPaso0 : BOOL;
    otraLuzPaso7 : BOOL;

    (* --- Resultados: 0 = pendiente, 1 = pasa, 2 = falla --- *)
    resultado : ARRAY[0..8] OF INT;
    nPasan    : INT;
    veredicto : INT := 0;
    i         : INT;
END_VAR

(* 1. Definicion del paso en curso *)
IF NOT finalizado THEN
    CASE paso OF
        0:  (* Reposo deshabilitado: V y R deben permanecer apagadas *)
            habilitado := FALSE; tEspera := T#200MS;
        1:  (* Al habilitar arranca en verde *)
            habilitado := TRUE;  tEspera := T#200MS;
            espV := TRUE;  espA := FALSE; espR := FALSE;

        (* --- Primer ciclo completo --- *)
        2:  (* 20 s de verde -> amarillo *)
            tEspera := T#20S;  espV := FALSE; espA := TRUE;  espR := FALSE;
        3:  (* 4 s de amarillo -> rojo *)
            tEspera := T#4S;   espV := FALSE; espA := FALSE; espR := TRUE;
        4:  (* 15 s de rojo -> verde *)
            tEspera := T#15S;  espV := TRUE;  espA := FALSE; espR := FALSE;

        (* --- Segundo ciclo: confirma que es ciclico y deja el semaforo en
               ROJO, que es la fase desde la que hay que interrumpir para que
               el reinicio en verde sea observable (enmienda 8) --- *)
        5:  (* 20 s de verde -> amarillo *)
            tEspera := T#20S;  espV := FALSE; espA := TRUE;  espR := FALSE;
        6:  (* 4 s de amarillo -> rojo *)
            tEspera := T#4S;   espV := FALSE; espA := FALSE; espR := TRUE;

        (* --- Intermitente e inhibicion --- *)
        7:  (* Se deshabilita ESTANDO EN ROJO: amarillo intermitente medido,
               con V y R vigiladas de forma continua *)
            habilitado := FALSE; tEspera := T#7S;
        8:  (* Al rehabilitar debe reiniciar EN VERDE, no continuar en rojo *)
            habilitado := TRUE;  tEspera := T#200MS;
            espV := TRUE;  espA := FALSE; espR := FALSE;
    END_CASE
END_IF

(* 2. Temporizadores del banco *)
tPaso(IN := NOT pulsoReset, PT := tEspera);
tCrono(IN := TRUE, PT := T_CRONO);
pulsoReset := FALSE;

(* 3. Llamada al bloque bajo prueba *)
fb(habilitado := habilitado);

(* 4. Medida de los intervalos del amarillo intermitente (paso 7).
      Duracion por diferencia de dos lecturas del cronometro libre. *)
IF paso = 7 THEN
    IF (fb.luzA AND NOT prevA) OR ((NOT fb.luzA) AND prevA) THEN
        IF primer THEN
            duracion := tCrono.ET - etFlanco;
            IF NOT fb.luzA THEN
                nOn := nOn + 1;
            ELSE
                nOff := nOff + 1;
            END_IF
            IF duracion < TOL_MIN OR duracion > TOL_MAX THEN
                error := TRUE;
            END_IF
        ELSE
            primer := TRUE;
        END_IF
        etFlanco := tCrono.ET;
    END_IF
END_IF
prevA := fb.luzA;

(* 5. Vigilancia continua y enclavada de las demas luces durante los pasos
      deshabilitados (enmienda 6). Un unico muestreo no sirve: si la
      implementacion alterna el amarillo con otra luz, la fase decide si se
      la sorprende encendida. *)
IF paso = 0 AND (fb.luzV OR fb.luzR) THEN
    otraLuzPaso0 := TRUE;
END_IF
IF paso = 7 AND (fb.luzV OR fb.luzR) THEN
    otraLuzPaso7 := TRUE;
END_IF

(* 6. Evaluacion al vencer el asentamiento del paso *)
IF tPaso.Q AND NOT finalizado THEN
    IF    (paso = 0 AND NOT fb.luzV AND NOT fb.luzR AND NOT otraLuzPaso0)
       OR (paso = 7 AND NOT fb.luzV AND NOT fb.luzR AND NOT otraLuzPaso7
                    AND nOn >= 2 AND nOff >= 2 AND NOT error)
       OR (paso <> 0 AND paso <> 7
                    AND fb.luzV = espV AND fb.luzA = espA AND fb.luzR = espR)
    THEN
        resultado[paso] := 1;
    ELSE
        resultado[paso] := 2;
    END_IF

    pulsoReset := TRUE;

    IF paso < ULTIMO_PASO THEN
        paso := paso + 1;
    ELSE
        finalizado := TRUE;
    END_IF
END_IF

(* 7. Veredicto global *)
IF finalizado AND veredicto = 0 THEN
    nPasan := 0;
    FOR i := 0 TO ULTIMO_PASO DO
        IF resultado[i] = 1 THEN
            nPasan := nPasan + 1;
        END_IF
    END_FOR

    IF nPasan = (ULTIMO_PASO + 1) THEN
        veredicto := 1;
    ELSE
        veredicto := 2;
    END_IF
END_IF
